Universal Robots URScript: FaiChun_9 Jan_10.script

def Machining1():
  # Default parameters:
  global speed_ms = 0.01
  global speed_rads = 0.75
  global accel_mss = 3
  global accel_radss = 1.2
  global blend_radius_m = 0.0003

  # Add subprograms here
  # Start of main program
  # Program generated by RoboDK v5.6.8 for UR10e on 10/01/2025 15:07:00
  # Using nominal kinematics.
  blend_radius_m = 0.0003
  speed_ms = 0.01
  # set_reference(p[0.340000, -0.015000, 0.001500, 0.000000, 0.000000, 0.000000])
  set_tcp(p[0.000000, 0.000000, 0.252000, 0.000000, 0.000000, 0.000000])
  # Show Tool
  movej([0.358985, -0.895332, -2.200270, -1.616787, 1.570796, 1.929781],accel_radss,speed_rads,0,blend_radius_m)
  movel([0.358985, -1.122148, -2.673539, -0.916702, 1.570796, 1.929781],accel_mss,speed_ms,0,blend_radius_m)
  #SetTool1
  #M_RunCode6
  #SetRPM60000
  speed_ms = 0.01
  #M_RunCode3
  movel([0.358985, -1.149717, -2.688845, -0.873826, 1.570796, 1.929781],accel_mss,speed_ms,0,blend_radius_m)
  speed_ms = 0.003
  movel([0.358985, -1.157003, -2.692612, -0.862774, 1.570796, 1.929781],accel_mss,speed_ms,0,blend_radius_m)
  speed_ms = 0.007
  movel([0.360284, -1.155838, -2.693115, -0.863435, 1.570796, 1.931080],accel_mss,speed_ms,0,blend_radius_m)
  movel([0.363800, -1.153166, -2.694264, -0.864959, 1.570796, 1.934596],accel_mss,speed_ms,0,blend_radius_m)
  movel([0.367667, -1.151137, -2.695132, -0.866120, 1.570796, 1.938463],accel_mss,speed_ms,0,blend_radius_m)
  movel([0.371673, -1.149666, -2.695758, -0.866965, 1.570796, 1.942469],accel_mss,speed_ms,0,blend_radius_m)
  movel([0.375593, -1.148672, -2.696180, -0.867537, 1.570796, 1.946389],accel_mss,speed_ms,0,blend_radius_m)
  movel([0.385811, -1.147094, -2.696848, -0.868447, 1.570796, 1.956607],accel_mss,speed_ms,0,blend_radius_m)
  movel([0.395233, -1.145814, -2.697388, -0.869187, 1.570796, 1.966029],accel_mss,speed_ms,0,blend_radius_m)
  movel([0.398878, -1.144990, -2.697734, -0.869664, 1.570796, 1.969674],accel_mss,speed_ms,0,blend_radius_m)
  movel([0.402533, -1.143763, -2.698250, -0.870377, 1.570796, 1.973330],accel_mss,speed_ms,0,blend_radius_m)
  movel([0.406011, -1.142059, -2.698963, -0.871368, 1.570796, 1.976808],accel_mss,speed_ms,0,blend_radius_m)
  movel([0.409148, -1.139796, -2.699904, -0.872688, 1.570796, 1.979944],accel_mss,speed_ms,0,blend_radius_m)
  movel([0.412438, -1.136413, -2.701304, -0.874672, 1.570796, 1.983234],accel_mss,speed_ms,0,blend_radius_m)
  movel([0.413570, -1.134739, -2.701992, -0.875658, 1.570796, 1.984366],accel_mss,speed_ms,0,blend_radius_m)
  movel([0.414360, -1.133075, -2.702674, -0.876641, 1.570796, 1.985156],accel_mss,speed_ms,0,blend_radius_m)
  movel([0.414991, -1.130073, -2.703896, -0.878420, 1.570796, 1.985787],accel_mss,speed_ms,0,blend_radius_m)
  movel([0.414425, -1.127699, -2.704856, -0.879834, 1.570796, 1.985221],accel_mss,speed_ms,0,blend_radius_m)
  movel([0.413477, -1.126577, -2.705309, -0.880504, 1.570796, 1.984274],accel_mss,speed_ms,0,blend_radius_m)
  movel([0.412318, -1.126143, -2.705483, -0.880763, 1.570796, 1.983114],accel_mss,speed_ms,0,blend_radius_m)
  movel([0.411061, -1.126342, -2.705403, -0.880644, 1.570796, 1.981857],accel_mss,speed_ms,0,blend_radius_m)
  movel([0.409841, -1.127103, -2.705097, -0.880189, 1.570796, 1.980638],accel_mss,speed_ms,0,blend_radius_m)
  movel([0.408484, -1.128982, -2.704338, -0.879069, 1.570796, 1.979281],accel_mss,speed_ms,0,blend_radius_m)
  movel([0.407268, -1.130867, -2.703573, -0.877948, 1.570796, 1.978064],accel_mss,speed_ms,0,blend_radius_m)
  movel([0.405338, -1.132846, -2.702767, -0.876776, 1.570796, 1.976135],accel_mss,speed_ms,0,blend_radius_m)
  movel([0.402737, -1.134615, -2.702043, -0.875731, 1.570796, 1.973533],accel_mss,speed_ms,0,blend_radius_m)
  movel([0.400364, -1.135207, -2.701800, -0.875382, 1.570796, 1.971160],accel_mss,speed_ms,0,blend_radius_m)
  movel([0.398406, -1.134766, -2.701981, -0.875642, 1.570796, 1.969202],accel_mss,speed_ms,0,blend_radius_m)
  movel([0.397035, -1.133442, -2.702523, -0.876424, 1.570796, 1.967832],accel_mss,speed_ms,0,blend_radius_m)
  movel([0.396404, -1.131466, -2.703330, -0.877593, 1.570796, 1.967200],accel_mss,speed_ms,0,blend_radius_m)
  movel([0.396662, -1.129077, -2.704300, -0.879013, 1.570796, 1.967458],accel_mss,speed_ms,0,blend_radius_m)
  movel([0.397874, -1.126522, -2.705330, -0.880536, 1.570796, 1.968671],accel_mss,speed_ms,0,blend_radius_m)
  movel([0.400111, -1.124058, -2.706319, -0.882012, 1.570796, 1.970908],accel_mss,speed_ms,0,blend_radius_m)
  movel([0.402368, -1.122361, -2.706996, -0.883031, 1.570796, 1.973164],accel_mss,speed_ms,0,blend_radius_m)
  movel([0.404592, -1.121272, -2.707430, -0.883687, 1.570796, 1.975389],accel_mss,speed_ms,0,blend_radius_m)
  movel([0.406779, -1.120798, -2.707618, -0.883973, 1.570796, 1.977575],accel_mss,speed_ms,0,blend_radius_m)
  movel([0.408920, -1.120940, -2.707561, -0.883887, 1.570796, 1.979716],accel_mss,speed_ms,0,blend_radius_m)
  movel([0.410941, -1.121627, -2.707288, -0.883473, 1.570796, 1.981737],accel_mss,speed_ms,0,blend_radius_m)
  movel([0.412761, -1.122788, -2.706826, -0.882775, 1.570796, 1.983557],accel_mss,speed_ms,0,blend_radius_m)
  movel([0.415800, -1.126514, -2.705334, -0.880541, 1.570796, 1.986596],accel_mss,speed_ms,0,blend_radius_m)
  movel([0.417144, -1.129442, -2.704152, -0.878795, 1.570796, 1.987940],accel_mss,speed_ms,0,blend_radius_m)
  movel([0.417974, -1.132572, -2.702879, -0.876938, 1.570796, 1.988771],accel_mss,speed_ms,0,blend_radius_m)
  movel([0.418302, -1.135897, -2.701516, -0.874976, 1.570796, 1.989099],accel_mss,speed_ms,0,blend_radius_m)
  movel([0.418128, -1.139411, -2.700064, -0.872914, 1.570796, 1.988924],accel_mss,speed_ms,0,blend_radius_m)
  movel([0.417267, -1.142978, -2.698578, -0.870833, 1.570796, 1.988063],accel_mss,speed_ms,0,blend_radius_m)
  movel([0.415537, -1.146458, -2.697116, -0.868815, 1.570796, 1.986334],accel_mss,speed_ms,0,blend_radius_m)
  movel([0.412946, -1.149856, -2.695677, -0.866856, 1.570796, 1.983742],accel_mss,speed_ms,0,blend_radius_m)
  movel([0.409498, -1.153176, -2.694260, -0.864954, 1.570796, 1.980294],accel_mss,speed_ms,0,blend_radius_m)
  movel([0.406063, -1.155728, -2.693163, -0.863498, 1.570796, 1.976860],accel_mss,speed_ms,0,blend_radius_m)
  movel([0.402585, -1.157607, -2.692351, -0.862431, 1.570796, 1.973381],accel_mss,speed_ms,0,blend_radius_m)
  movel([0.399151, -1.158929, -2.691777, -0.861683, 1.570796, 1.969948],accel_mss,speed_ms,0,blend_radius_m)
  movel([0.395859, -1.159805, -2.691396, -0.861188, 1.570796, 1.966655],accel_mss,speed_ms,0,blend_radius_m)
  movel([0.388031, -1.160961, -2.690892, -0.860535, 1.570796, 1.958827],accel_mss,speed_ms,0,blend_radius_m)
  movel([0.380613, -1.162143, -2.690376, -0.859870, 1.570796, 1.951410],accel_mss,speed_ms,0,blend_radius_m)
  movel([0.377615, -1.162965, -2.690015, -0.859408, 1.570796, 1.948411],accel_mss,speed_ms,0,blend_radius_m)
  movel([0.374545, -1.164177, -2.689483, -0.858729, 1.570796, 1.945341],accel_mss,speed_ms,0,blend_radius_m)
  movel([0.371509, -1.165851, -2.688746, -0.857792, 1.570796, 1.942306],accel_mss,speed_ms,0,blend_radius_m)
  movel([0.368622, -1.168057, -2.687769, -0.856563, 1.570796, 1.939418],accel_mss,speed_ms,0,blend_radius_m)
  movel([0.369262, -1.169016, -2.687343, -0.856030, 1.570796, 1.940058],accel_mss,speed_ms,0,blend_radius_m)
  movel([0.371229, -1.171492, -2.686239, -0.854659, 1.570796, 1.942025],accel_mss,speed_ms,0,blend_radius_m)
  movel([0.373363, -1.173304, -2.685426, -0.853659, 1.570796, 1.944159],accel_mss,speed_ms,0,blend_radius_m)
  movel([0.375672, -1.174449, -2.684911, -0.853029, 1.570796, 1.946468],accel_mss,speed_ms,0,blend_radius_m)
  movel([0.378153, -1.174934, -2.684692, -0.852763, 1.570796, 1.948949],accel_mss,speed_ms,0,blend_radius_m)
  movel([0.380756, -1.174836, -2.684736, -0.852816, 1.570796, 1.951553],accel_mss,speed_ms,0,blend_radius_m)
  movel([0.383422, -1.174230, -2.685010, -0.853150, 1.570796, 1.954218],accel_mss,speed_ms,0,blend_radius_m)
  movel([0.386160, -1.173110, -2.685513, -0.853766, 1.570796, 1.956957],accel_mss,speed_ms,0,blend_radius_m)
  movel([0.388972, -1.171476, -2.686246, -0.854667, 1.570796, 1.959768],accel_mss,speed_ms,0,blend_radius_m)
  movel([0.376141, -1.182465, -2.681266, -0.848658, 1.570796, 1.946938],accel_mss,speed_ms,0,blend_radius_m)
  movel([0.358985, -1.157003, -2.692612, -0.862774, 1.570796, 1.929781],accel_mss,speed_ms,0,blend_radius_m)
  speed_ms = 0.003
  movel([0.358985, -1.149717, -2.688845, -0.873826, 1.570796, 1.929781],accel_mss,speed_ms,0,blend_radius_m)
  speed_ms = 0.01
  movel([0.358985, -1.122148, -2.673539, -0.916702, 1.570796, 1.929781],accel_mss,speed_ms,0,blend_radius_m)
  #M_RunCode9
  movel([0.390070, -1.155228, -2.659313, -0.897848, 1.570796, 1.960867],accel_mss,speed_ms,0,blend_radius_m)
  #M_RunCode3
  movel([0.390070, -1.182636, -2.674188, -0.855565, 1.570796, 1.960867],accel_mss,speed_ms,0,blend_radius_m)
  speed_ms = 0.003
  movel([0.390070, -1.189858, -2.677844, -0.844687, 1.570796, 1.960867],accel_mss,speed_ms,0,blend_radius_m)
  speed_ms = 0.007
  movel([0.396700, -1.183388, -2.680842, -0.848159, 1.570796, 1.967497],accel_mss,speed_ms,0,blend_radius_m)
  movel([0.406631, -1.174785, -2.684760, -0.852845, 1.570796, 1.977428],accel_mss,speed_ms,0,blend_radius_m)
  movel([0.416940, -1.166524, -2.688448, -0.857416, 1.570796, 1.987736],accel_mss,speed_ms,0,blend_radius_m)
  movel([0.424558, -1.161153, -2.690809, -0.860427, 1.570796, 1.995354],accel_mss,speed_ms,0,blend_radius_m)
  movel([0.427380, -1.159602, -2.691485, -0.861302, 1.570796, 1.998176],accel_mss,speed_ms,0,blend_radius_m)
  movel([0.429592, -1.158857, -2.691809, -0.861723, 1.570796, 2.000389],accel_mss,speed_ms,0,blend_radius_m)
  movel([0.431192, -1.158925, -2.691779, -0.861685, 1.570796, 2.001988],accel_mss,speed_ms,0,blend_radius_m)
  movel([0.432177, -1.159797, -2.691400, -0.861192, 1.570796, 2.002973],accel_mss,speed_ms,0,blend_radius_m)
  movel([0.432434, -1.161264, -2.690760, -0.860365, 1.570796, 2.003230],accel_mss,speed_ms,0,blend_radius_m)
  movel([0.431856, -1.163109, -2.689953, -0.859328, 1.570796, 2.002653],accel_mss,speed_ms,0,blend_radius_m)
  movel([0.430453, -1.165326, -2.688977, -0.858086, 1.570796, 2.001249],accel_mss,speed_ms,0,blend_radius_m)
  movel([0.428224, -1.167916, -2.687832, -0.856641, 1.570796, 1.999021],accel_mss,speed_ms,0,blend_radius_m)
  movel([0.421358, -1.174456, -2.684908, -0.853025, 1.570796, 1.992155],accel_mss,speed_ms,0,blend_radius_m)
  movel([0.411361, -1.182965, -2.681036, -0.848388, 1.570796, 1.982158],accel_mss,speed_ms,0,blend_radius_m)
  movel([0.401263, -1.190989, -2.677315, -0.844085, 1.570796, 1.972059],accel_mss,speed_ms,0,blend_radius_m)
  movel([0.393942, -1.196149, -2.674885, -0.841355, 1.570796, 1.964739],accel_mss,speed_ms,0,blend_radius_m)
  movel([0.391243, -1.197643, -2.674176, -0.840570, 1.570796, 1.962040],accel_mss,speed_ms,0,blend_radius_m)
  movel([0.389113, -1.198381, -2.673825, -0.840183, 1.570796, 1.959910],accel_mss,speed_ms,0,blend_radius_m)
  movel([0.387547, -1.198358, -2.673836, -0.840195, 1.570796, 1.958343],accel_mss,speed_ms,0,blend_radius_m)
  movel([0.386539, -1.197580, -2.674206, -0.840603, 1.570796, 1.957335],accel_mss,speed_ms,0,blend_radius_m)
  movel([0.386213, -1.196230, -2.674847, -0.841312, 1.570796, 1.957009],accel_mss,speed_ms,0,blend_radius_m)
  movel([0.386687, -1.194496, -2.675667, -0.842226, 1.570796, 1.957483],accel_mss,speed_ms,0,blend_radius_m)
  movel([0.387972, -1.192374, -2.676665, -0.843349, 1.570796, 1.958769],accel_mss,speed_ms,0,blend_radius_m)
  movel([0.390070, -1.189858, -2.677844, -0.844687, 1.570796, 1.960867],accel_mss,speed_ms,0,blend_radius_m)
  speed_ms = 0.003
  movel([0.390070, -1.182636, -2.674188, -0.855565, 1.570796, 1.960867],accel_mss,speed_ms,0,blend_radius_m)
  speed_ms = 0.01
  movel([0.390070, -1.155228, -2.659313, -0.897848, 1.570796, 1.960867],accel_mss,speed_ms,0,blend_radius_m)
  #M_RunCode9
  movel([0.383757, -1.157911, -2.658112, -0.896367, 1.570796, 1.954554],accel_mss,speed_ms,0,blend_radius_m)
  #M_RunCode3
  movel([0.383757, -1.185302, -2.672951, -0.854136, 1.570796, 1.954554],accel_mss,speed_ms,0,blend_radius_m)
  speed_ms = 0.003
  movel([0.383757, -1.192518, -2.676598, -0.843273, 1.570796, 1.954554],accel_mss,speed_ms,0,blend_radius_m)
  speed_ms = 0.007
  movel([0.384034, -1.190067, -2.677746, -0.844576, 1.570796, 1.954830],accel_mss,speed_ms,0,blend_radius_m)
  movel([0.384719, -1.187441, -2.678969, -0.845979, 1.570796, 1.955516],accel_mss,speed_ms,0,blend_radius_m)
  movel([0.385830, -1.184674, -2.680249, -0.847465, 1.570796, 1.956626],accel_mss,speed_ms,0,blend_radius_m)
  movel([0.387369, -1.181762, -2.681588, -0.849039, 1.570796, 1.958165],accel_mss,speed_ms,0,blend_radius_m)
  movel([0.389339, -1.178702, -2.682986, -0.850702, 1.570796, 1.960136],accel_mss,speed_ms,0,blend_radius_m)
  movel([0.391735, -1.175551, -2.684414, -0.852424, 1.570796, 1.962531],accel_mss,speed_ms,0,blend_radius_m)
  movel([0.394540, -1.172369, -2.685846, -0.854174, 1.570796, 1.965337],accel_mss,speed_ms,0,blend_radius_m)
  movel([0.397760, -1.169157, -2.687280, -0.855952, 1.570796, 1.968556],accel_mss,speed_ms,0,blend_radius_m)
  movel([0.401398, -1.165917, -2.688716, -0.857755, 1.570796, 1.972194],accel_mss,speed_ms,0,blend_radius_m)
  movel([0.405183, -1.162881, -2.690052, -0.859456, 1.570796, 1.975979],accel_mss,speed_ms,0,blend_radius_m)
  movel([0.408839, -1.160283, -2.691188, -0.860918, 1.570796, 1.979636],accel_mss,speed_ms,0,blend_radius_m)
  movel([0.412361, -1.158134, -2.692122, -0.862133, 1.570796, 1.983157],accel_mss,speed_ms,0,blend_radius_m)
  movel([0.415741, -1.156438, -2.692856, -0.863094, 1.570796, 1.986537],accel_mss,speed_ms,0,blend_radius_m)
  movel([0.418920, -1.155194, -2.693393, -0.863802, 1.570796, 1.989717],accel_mss,speed_ms,0,blend_radius_m)
  movel([0.421843, -1.154407, -2.693731, -0.864250, 1.570796, 1.992639],accel_mss,speed_ms,0,blend_radius_m)
  movel([0.424499, -1.154076, -2.693874, -0.864439, 1.570796, 1.995295],accel_mss,speed_ms,0,blend_radius_m)
  movel([0.426890, -1.154203, -2.693819, -0.864367, 1.570796, 1.997687],accel_mss,speed_ms,0,blend_radius_m)
  movel([0.428991, -1.154756, -2.693581, -0.864051, 1.570796, 1.999787],accel_mss,speed_ms,0,blend_radius_m)
  movel([0.430782, -1.155707, -2.693172, -0.863511, 1.570796, 2.001578],accel_mss,speed_ms,0,blend_radius_m)
  movel([0.432260, -1.157045, -2.692594, -0.862750, 1.570796, 2.003056],accel_mss,speed_ms,0,blend_radius_m)
  movel([0.433430, -1.158771, -2.691846, -0.861772, 1.570796, 2.004226],accel_mss,speed_ms,0,blend_radius_m)
  movel([0.434237, -1.160788, -2.690968, -0.860633, 1.570796, 2.005033],accel_mss,speed_ms,0,blend_radius_m)
  movel([0.434638, -1.162993, -2.690003, -0.859393, 1.570796, 2.005434],accel_mss,speed_ms,0,blend_radius_m)
  movel([0.434635, -1.165385, -2.688951, -0.858052, 1.570796, 2.005431],accel_mss,speed_ms,0,blend_radius_m)
  movel([0.434233, -1.167961, -2.687812, -0.856616, 1.570796, 2.005030],accel_mss,speed_ms,0,blend_radius_m)
  movel([0.433415, -1.170685, -2.686599, -0.855105, 1.570796, 2.004211],accel_mss,speed_ms,0,blend_radius_m)
  movel([0.432178, -1.173518, -2.685330, -0.853541, 1.570796, 2.002974],accel_mss,speed_ms,0,blend_radius_m)
  movel([0.430522, -1.176455, -2.684005, -0.851929, 1.570796, 2.001318],accel_mss,speed_ms,0,blend_radius_m)
  movel([0.428448, -1.179502, -2.682621, -0.850266, 1.570796, 1.999245],accel_mss,speed_ms,0,blend_radius_m)
  movel([0.425982, -1.182592, -2.681208, -0.848589, 1.570796, 1.996779],accel_mss,speed_ms,0,blend_radius_m)
  movel([0.423147, -1.185664, -2.679792, -0.846933, 1.570796, 1.993943],accel_mss,speed_ms,0,blend_radius_m)
  movel([0.419941, -1.188728, -2.678370, -0.845290, 1.570796, 1.990737],accel_mss,speed_ms,0,blend_radius_m)
  movel([0.416367, -1.191779, -2.676945, -0.843665, 1.570796, 1.987163],accel_mss,speed_ms,0,blend_radius_m)
  movel([0.412690, -1.194608, -2.675614, -0.842167, 1.570796, 1.983486],accel_mss,speed_ms,0,blend_radius_m)
  movel([0.409169, -1.197005, -2.674479, -0.840905, 1.570796, 1.979965],accel_mss,speed_ms,0,blend_radius_m)
  movel([0.405805, -1.198977, -2.673541, -0.839871, 1.570796, 1.976601],accel_mss,speed_ms,0,blend_radius_m)
  movel([0.402584, -1.200530, -2.672799, -0.839060, 1.570796, 1.973380],accel_mss,speed_ms,0,blend_radius_m)
  movel([0.399556, -1.201668, -2.672254, -0.838467, 1.570796, 1.970353],accel_mss,speed_ms,0,blend_radius_m)
  movel([0.396767, -1.202400, -2.671902, -0.838087, 1.570796, 1.967564],accel_mss,speed_ms,0,blend_radius_m)
  movel([0.394210, -1.202727, -2.671745, -0.837916, 1.570796, 1.965007],accel_mss,speed_ms,0,blend_radius_m)
  movel([0.391887, -1.202647, -2.671784, -0.837958, 1.570796, 1.962683],accel_mss,speed_ms,0,blend_radius_m)
  movel([0.389820, -1.202186, -2.672006, -0.838198, 1.570796, 1.960616],accel_mss,speed_ms,0,blend_radius_m)
  movel([0.388028, -1.201364, -2.672400, -0.838625, 1.570796, 1.958824],accel_mss,speed_ms,0,blend_radius_m)
  movel([0.386519, -1.200177, -2.672968, -0.839244, 1.570796, 1.957315],accel_mss,speed_ms,0,blend_radius_m)
  movel([0.385286, -1.198629, -2.673707, -0.840053, 1.570796, 1.956082],accel_mss,speed_ms,0,blend_radius_m)
  movel([0.384388, -1.196795, -2.674579, -0.841015, 1.570796, 1.955184],accel_mss,speed_ms,0,blend_radius_m)
  movel([0.383876, -1.194758, -2.675543, -0.842088, 1.570796, 1.954672],accel_mss,speed_ms,0,blend_radius_m)
  movel([0.383757, -1.192518, -2.676598, -0.843273, 1.570796, 1.954554],accel_mss,speed_ms,0,blend_radius_m)
  speed_ms = 0.003
  movel([0.383757, -1.185302, -2.672951, -0.854136, 1.570796, 1.954554],accel_mss,speed_ms,0,blend_radius_m)
  speed_ms = 0.01
  movel([0.383757, -1.157911, -2.658112, -0.896367, 1.570796, 1.954554],accel_mss,speed_ms,0,blend_radius_m)
  #M_RunCode9
  movel([0.496093, -1.382466, -2.528375, -0.801548, 1.570796, 2.066889],accel_mss,speed_ms,0,blend_radius_m)
  #M_RunCode3
  movel([0.496093, -1.406789, -2.540293, -0.765307, 1.570796, 2.066889],accel_mss,speed_ms,0,blend_radius_m)
  speed_ms = 0.003
  movel([0.496093, -1.413093, -2.543201, -0.756095, 1.570796, 2.066889],accel_mss,speed_ms,0,blend_radius_m)
  speed_ms = 0.007
  movel([0.497104, -1.412495, -2.543652, -0.756242, 1.570796, 2.067901],accel_mss,speed_ms,0,blend_radius_m)
  movel([0.499783, -1.411227, -2.544607, -0.756556, 1.570796, 2.070579],accel_mss,speed_ms,0,blend_radius_m)
  movel([0.502622, -1.410494, -2.545157, -0.756738, 1.570796, 2.073418],accel_mss,speed_ms,0,blend_radius_m)
  movel([0.505487, -1.410196, -2.545381, -0.756812, 1.570796, 2.076283],accel_mss,speed_ms,0,blend_radius_m)
  movel([0.508237, -1.410226, -2.545358, -0.756805, 1.570796, 2.079034],accel_mss,speed_ms,0,blend_radius_m)
  movel([0.515289, -1.411028, -2.544756, -0.756605, 1.570796, 2.086086],accel_mss,speed_ms,0,blend_radius_m)
  movel([0.521765, -1.411881, -2.544115, -0.756394, 1.570796, 2.092561],accel_mss,speed_ms,0,blend_radius_m)
  movel([0.524304, -1.411969, -2.544048, -0.756372, 1.570796, 2.095101],accel_mss,speed_ms,0,blend_radius_m)
  movel([0.526887, -1.411770, -2.544198, -0.756421, 1.570796, 2.097684],accel_mss,speed_ms,0,blend_radius_m)
  movel([0.529402, -1.411199, -2.544627, -0.756563, 1.570796, 2.100198],accel_mss,speed_ms,0,blend_radius_m)
  movel([0.531734, -1.410169, -2.545401, -0.756819, 1.570796, 2.102530],accel_mss,speed_ms,0,blend_radius_m)
  movel([0.534284, -1.408370, -2.546748, -0.757271, 1.570796, 2.105081],accel_mss,speed_ms,0,blend_radius_m)
  movel([0.535210, -1.407391, -2.547480, -0.757519, 1.570796, 2.106007],accel_mss,speed_ms,0,blend_radius_m)
  movel([0.535902, -1.406358, -2.548250, -0.757782, 1.570796, 2.106698],accel_mss,speed_ms,0,blend_radius_m)
  movel([0.536626, -1.404345, -2.549745, -0.758299, 1.570796, 2.107423],accel_mss,speed_ms,0,blend_radius_m)
  movel([0.536483, -1.402557, -2.551069, -0.758763, 1.570796, 2.107279],accel_mss,speed_ms,0,blend_radius_m)
  movel([0.535964, -1.401585, -2.551787, -0.759017, 1.570796, 2.106761],accel_mss,speed_ms,0,blend_radius_m)
  movel([0.535230, -1.401062, -2.552172, -0.759155, 1.570796, 2.106027],accel_mss,speed_ms,0,blend_radius_m)
  movel([0.534373, -1.400967, -2.552242, -0.759180, 1.570796, 2.105170],accel_mss,speed_ms,0,blend_radius_m)
  movel([0.533483, -1.401277, -2.552014, -0.759098, 1.570796, 2.104279],accel_mss,speed_ms,0,blend_radius_m)
  movel([0.532384, -1.402355, -2.551218, -0.758816, 1.570796, 2.103180],accel_mss,speed_ms,0,blend_radius_m)
  movel([0.531379, -1.403465, -2.550397, -0.758527, 1.570796, 2.102176],accel_mss,speed_ms,0,blend_radius_m)
  movel([0.529890, -1.404508, -2.549624, -0.758257, 1.570796, 2.100686],accel_mss,speed_ms,0,blend_radius_m)
  movel([0.527963, -1.405280, -2.549051, -0.758058, 1.570796, 2.098760],accel_mss,speed_ms,0,blend_radius_m)
  movel([0.526316, -1.405254, -2.549070, -0.758064, 1.570796, 2.097112],accel_mss,speed_ms,0,blend_radius_m)
  movel([0.525050, -1.404571, -2.549577, -0.758240, 1.570796, 2.095846],accel_mss,speed_ms,0,blend_radius_m)
  movel([0.524270, -1.403366, -2.550470, -0.758552, 1.570796, 2.095067],accel_mss,speed_ms,0,blend_radius_m)
  movel([0.524055, -1.401836, -2.551601, -0.758951, 1.570796, 2.094851],accel_mss,speed_ms,0,blend_radius_m)
  movel([0.524478, -1.400181, -2.552821, -0.759387, 1.570796, 2.095274],accel_mss,speed_ms,0,blend_radius_m)
  movel([0.525555, -1.398592, -2.553988, -0.759809, 1.570796, 2.096352],accel_mss,speed_ms,0,blend_radius_m)
  movel([0.527302, -1.397266, -2.554959, -0.760164, 1.570796, 2.098099],accel_mss,speed_ms,0,blend_radius_m)
  movel([0.528984, -1.396492, -2.555524, -0.760372, 1.570796, 2.099781],accel_mss,speed_ms,0,blend_radius_m)
  movel([0.530578, -1.396145, -2.555778, -0.760466, 1.570796, 2.101374],accel_mss,speed_ms,0,blend_radius_m)
  movel([0.532081, -1.396224, -2.555720, -0.760445, 1.570796, 2.102877],accel_mss,speed_ms,0,blend_radius_m)
  movel([0.533493, -1.396734, -2.555347, -0.760307, 1.570796, 2.104290],accel_mss,speed_ms,0,blend_radius_m)
  movel([0.534769, -1.397605, -2.554711, -0.760073, 1.570796, 2.105566],accel_mss,speed_ms,0,blend_radius_m)
  movel([0.535865, -1.398770, -2.553857, -0.759762, 1.570796, 2.106661],accel_mss,speed_ms,0,blend_radius_m)
  movel([0.537521, -1.401976, -2.551498, -0.758915, 1.570796, 2.108317],accel_mss,speed_ms,0,blend_radius_m)
  movel([0.538126, -1.404299, -2.549779, -0.758311, 1.570796, 2.108923],accel_mss,speed_ms,0,blend_radius_m)
  movel([0.538374, -1.406672, -2.548015, -0.757702, 1.570796, 2.109170],accel_mss,speed_ms,0,blend_radius_m)
  movel([0.538264, -1.409089, -2.546211, -0.757090, 1.570796, 2.109060],accel_mss,speed_ms,0,blend_radius_m)
  movel([0.537801, -1.411550, -2.544364, -0.756476, 1.570796, 2.108597],accel_mss,speed_ms,0,blend_radius_m)
  movel([0.536875, -1.413924, -2.542573, -0.755892, 1.570796, 2.107671],accel_mss,speed_ms,0,blend_radius_m)
  movel([0.535368, -1.416086, -2.540936, -0.755367, 1.570796, 2.106164],accel_mss,speed_ms,0,blend_radius_m)
  movel([0.533284, -1.418039, -2.539451, -0.754899, 1.570796, 2.104080],accel_mss,speed_ms,0,blend_radius_m)
  movel([0.530625, -1.419784, -2.538119, -0.754486, 1.570796, 2.101421],accel_mss,speed_ms,0,blend_radius_m)
  movel([0.528047, -1.420988, -2.537198, -0.754204, 1.570796, 2.098844],accel_mss,speed_ms,0,blend_radius_m)
  movel([0.525504, -1.421702, -2.536650, -0.754037, 1.570796, 2.096300],accel_mss,speed_ms,0,blend_radius_m)
  movel([0.523046, -1.422024, -2.536403, -0.753962, 1.570796, 2.093842],accel_mss,speed_ms,0,blend_radius_m)
  movel([0.520727, -1.422052, -2.536382, -0.753956, 1.570796, 2.091523],accel_mss,speed_ms,0,blend_radius_m)
  movel([0.515303, -1.421445, -2.536847, -0.754097, 1.570796, 2.086099],accel_mss,speed_ms,0,blend_radius_m)
  movel([0.510152, -1.420924, -2.537247, -0.754219, 1.570796, 2.080948],accel_mss,speed_ms,0,blend_radius_m)
  movel([0.508029, -1.420964, -2.537216, -0.754209, 1.570796, 2.078825],accel_mss,speed_ms,0,blend_radius_m)
  movel([0.505817, -1.421270, -2.536982, -0.754138, 1.570796, 2.076613],accel_mss,speed_ms,0,blend_radius_m)
  movel([0.503574, -1.421917, -2.536485, -0.753987, 1.570796, 2.074370],accel_mss,speed_ms,0,blend_radius_m)
  movel([0.501367, -1.422986, -2.535664, -0.753740, 1.570796, 2.072163],accel_mss,speed_ms,0,blend_radius_m)
  movel([0.501695, -1.423803, -2.535035, -0.753552, 1.570796, 2.072492],accel_mss,speed_ms,0,blend_radius_m)
  movel([0.502756, -1.425977, -2.533355, -0.753056, 1.570796, 2.073552],accel_mss,speed_ms,0,blend_radius_m)
  movel([0.504008, -1.427693, -2.532026, -0.752670, 1.570796, 2.074805],accel_mss,speed_ms,0,blend_radius_m)
  movel([0.505454, -1.428956, -2.531044, -0.752389, 1.570796, 2.076250],accel_mss,speed_ms,0,blend_radius_m)
  movel([0.507091, -1.429766, -2.530413, -0.752210, 1.570796, 2.077887],accel_mss,speed_ms,0,blend_radius_m)
  movel([0.508876, -1.430170, -2.530098, -0.752121, 1.570796, 2.079672],accel_mss,speed_ms,0,blend_radius_m)
  movel([0.510757, -1.430216, -2.530063, -0.752111, 1.570796, 2.081553],accel_mss,speed_ms,0,blend_radius_m)
  movel([0.512740, -1.429904, -2.530306, -0.752179, 1.570796, 2.083536],accel_mss,speed_ms,0,blend_radius_m)
  movel([0.514827, -1.429230, -2.530831, -0.752328, 1.570796, 2.085623],accel_mss,speed_ms,0,blend_radius_m)
  movel([0.504898, -1.434894, -2.526397, -0.751098, 1.570796, 2.075694],accel_mss,speed_ms,0,blend_radius_m)
  movel([0.496093, -1.413093, -2.543201, -0.756095, 1.570796, 2.066889],accel_mss,speed_ms,0,blend_radius_m)
  speed_ms = 0.003
  movel([0.496093, -1.406789, -2.540293, -0.765307, 1.570796, 2.066889],accel_mss,speed_ms,0,blend_radius_m)
  speed_ms = 0.01
  movel([0.496093, -1.382466, -2.528375, -0.801548, 1.570796, 2.066889],accel_mss,speed_ms,0,blend_radius_m)
  #M_RunCode9
  movel([0.512138, -1.403973, -2.512554, -0.795862, 1.570796, 2.082934],accel_mss,speed_ms,0,blend_radius_m)
  #M_RunCode3
  movel([0.512138, -1.427879, -2.524206, -0.760304, 1.570796, 2.082934],accel_mss,speed_ms,0,blend_radius_m)
  speed_ms = 0.003
  movel([0.512138, -1.434068, -2.527046, -0.751275, 1.570796, 2.082934],accel_mss,speed_ms,0,blend_radius_m)
  speed_ms = 0.007
  movel([0.514003, -1.433320, -2.527634, -0.751435, 1.570796, 2.084799],accel_mss,speed_ms,0,blend_radius_m)
  movel([0.515626, -1.433332, -2.527624, -0.751432, 1.570796, 2.086422],accel_mss,speed_ms,0,blend_radius_m)
  movel([0.516887, -1.433975, -2.527119, -0.751294, 1.570796, 2.087684],accel_mss,speed_ms,0,blend_radius_m)
  movel([0.517657, -1.435128, -2.526212, -0.751048, 1.570796, 2.088453],accel_mss,speed_ms,0,blend_radius_m)
  movel([0.517868, -1.436594, -2.525056, -0.750738, 1.570796, 2.088665],accel_mss,speed_ms,0,blend_radius_m)
  movel([0.517453, -1.438175, -2.523806, -0.750408, 1.570796, 2.088249],accel_mss,speed_ms,0,blend_radius_m)
  movel([0.516413, -1.439679, -2.522613, -0.750097, 1.570796, 2.087209],accel_mss,speed_ms,0,blend_radius_m)
  movel([0.514754, -1.440917, -2.521629, -0.749844, 1.570796, 2.085550],accel_mss,speed_ms,0,blend_radius_m)
  movel([0.513217, -1.441589, -2.521093, -0.749707, 1.570796, 2.084014],accel_mss,speed_ms,0,blend_radius_m)
  movel([0.511950, -1.441787, -2.520935, -0.749667, 1.570796, 2.082746],accel_mss,speed_ms,0,blend_radius_m)
  movel([0.510647, -1.442088, -2.520695, -0.749606, 1.570796, 2.081443],accel_mss,speed_ms,0,blend_radius_m)
  movel([0.509919, -1.442689, -2.520215, -0.749485, 1.570796, 2.080715],accel_mss,speed_ms,0,blend_radius_m)
  movel([0.509449, -1.443526, -2.519546, -0.749317, 1.570796, 2.080245],accel_mss,speed_ms,0,blend_radius_m)
  movel([0.509278, -1.444452, -2.518804, -0.749133, 1.570796, 2.080074],accel_mss,speed_ms,0,blend_radius_m)
  movel([0.509440, -1.445324, -2.518105, -0.748960, 1.570796, 2.080236],accel_mss,speed_ms,0,blend_radius_m)
  movel([0.509993, -1.446284, -2.517333, -0.748772, 1.570796, 2.080789],accel_mss,speed_ms,0,blend_radius_m)
  movel([0.510801, -1.446988, -2.516767, -0.748634, 1.570796, 2.081597],accel_mss,speed_ms,0,blend_radius_m)
  movel([0.511865, -1.447436, -2.516405, -0.748547, 1.570796, 2.082661],accel_mss,speed_ms,0,blend_radius_m)
  movel([0.513186, -1.447631, -2.516249, -0.748510, 1.570796, 2.083982],accel_mss,speed_ms,0,blend_radius_m)
  movel([0.514688, -1.447559, -2.516306, -0.748524, 1.570796, 2.085484],accel_mss,speed_ms,0,blend_radius_m)
  movel([0.516291, -1.447213, -2.516585, -0.748591, 1.570796, 2.087087],accel_mss,speed_ms,0,blend_radius_m)
  movel([0.517999, -1.446591, -2.517086, -0.748712, 1.570796, 2.088795],accel_mss,speed_ms,0,blend_radius_m)
  movel([0.519813, -1.445693, -2.517809, -0.748888, 1.570796, 2.090609],accel_mss,speed_ms,0,blend_radius_m)
  movel([0.522666, -1.443719, -2.519391, -0.749279, 1.570796, 2.093462],accel_mss,speed_ms,0,blend_radius_m)
  movel([0.524983, -1.441258, -2.521357, -0.749774, 1.570796, 2.095780],accel_mss,speed_ms,0,blend_radius_m)
  movel([0.525915, -1.439851, -2.522477, -0.750062, 1.570796, 2.096711],accel_mss,speed_ms,0,blend_radius_m)
  movel([0.526652, -1.438341, -2.523675, -0.750373, 1.570796, 2.097449],accel_mss,speed_ms,0,blend_radius_m)
  movel([0.527554, -1.435008, -2.526307, -0.751074, 1.570796, 2.098351],accel_mss,speed_ms,0,blend_radius_m)
  movel([0.527587, -1.431347, -2.529179, -0.751863, 1.570796, 2.098383],accel_mss,speed_ms,0,blend_radius_m)
  movel([0.526637, -1.427456, -2.532210, -0.752723, 1.570796, 2.097433],accel_mss,speed_ms,0,blend_radius_m)
  movel([0.542111, -1.418898, -2.538796, -0.754695, 1.570796, 2.112907],accel_mss,speed_ms,0,blend_radius_m)
  movel([0.547688, -1.435758, -2.525716, -0.750915, 1.570796, 2.118485],accel_mss,speed_ms,0,blend_radius_m)
  movel([0.537746, -1.441111, -2.521474, -0.749804, 1.570796, 2.108543],accel_mss,speed_ms,0,blend_radius_m)
  movel([0.539901, -1.439199, -2.522994, -0.750196, 1.570796, 2.110697],accel_mss,speed_ms,0,blend_radius_m)
  movel([0.541670, -1.436872, -2.524837, -0.750680, 1.570796, 2.112466],accel_mss,speed_ms,0,blend_radius_m)
  movel([0.542959, -1.434240, -2.526912, -0.751238, 1.570796, 2.113756],accel_mss,speed_ms,0,blend_radius_m)
  movel([0.543680, -1.431418, -2.529124, -0.751847, 1.570796, 2.114477],accel_mss,speed_ms,0,blend_radius_m)
  movel([0.543769, -1.428514, -2.531388, -0.752487, 1.570796, 2.114565],accel_mss,speed_ms,0,blend_radius_m)
  movel([0.543166, -1.425645, -2.533613, -0.753131, 1.570796, 2.113962],accel_mss,speed_ms,0,blend_radius_m)
  movel([0.531802, -1.431868, -2.528772, -0.751749, 1.570796, 2.102598],accel_mss,speed_ms,0,blend_radius_m)
  movel([0.532645, -1.435321, -2.526060, -0.751007, 1.570796, 2.103441],accel_mss,speed_ms,0,blend_radius_m)
  movel([0.532812, -1.438966, -2.523179, -0.750244, 1.570796, 2.103608],accel_mss,speed_ms,0,blend_radius_m)
  movel([0.532201, -1.442603, -2.520284, -0.749502, 1.570796, 2.102997],accel_mss,speed_ms,0,blend_radius_m)
  movel([0.531565, -1.444346, -2.518889, -0.749154, 1.570796, 2.102361],accel_mss,speed_ms,0,blend_radius_m)
  movel([0.530709, -1.446043, -2.517527, -0.748819, 1.570796, 2.101506],accel_mss,speed_ms,0,blend_radius_m)
  movel([0.529618, -1.447639, -2.516242, -0.748508, 1.570796, 2.100414],accel_mss,speed_ms,0,blend_radius_m)
  movel([0.528273, -1.449088, -2.515072, -0.748229, 1.570796, 2.099070],accel_mss,speed_ms,0,blend_radius_m)
  movel([0.526675, -1.450389, -2.514018, -0.747982, 1.570796, 2.097472],accel_mss,speed_ms,0,blend_radius_m)
  movel([0.524823, -1.451546, -2.513080, -0.747764, 1.570796, 2.095619],accel_mss,speed_ms,0,blend_radius_m)
  movel([0.522889, -1.452474, -2.512325, -0.747590, 1.570796, 2.093685],accel_mss,speed_ms,0,blend_radius_m)
  movel([0.521038, -1.453096, -2.511818, -0.747475, 1.570796, 2.091834],accel_mss,speed_ms,0,blend_radius_m)
  movel([0.519270, -1.453408, -2.511564, -0.747417, 1.570796, 2.090067],accel_mss,speed_ms,0,blend_radius_m)
  movel([0.517584, -1.453415, -2.511558, -0.747416, 1.570796, 2.088380],accel_mss,speed_ms,0,blend_radius_m)
  movel([0.514548, -1.452701, -2.512140, -0.747548, 1.570796, 2.085344],accel_mss,speed_ms,0,blend_radius_m)
  movel([0.512020, -1.451143, -2.513407, -0.747839, 1.570796, 2.082816],accel_mss,speed_ms,0,blend_radius_m)
  movel([0.510039, -1.448945, -2.515187, -0.748257, 1.570796, 2.080835],accel_mss,speed_ms,0,blend_radius_m)
  movel([0.508638, -1.446319, -2.517305, -0.748765, 1.570796, 2.079434],accel_mss,speed_ms,0,blend_radius_m)
  movel([0.508085, -1.444283, -2.518939, -0.749166, 1.570796, 2.078881],accel_mss,speed_ms,0,blend_radius_m)
  movel([0.507919, -1.441997, -2.520768, -0.749624, 1.570796, 2.078716],accel_mss,speed_ms,0,blend_radius_m)
  movel([0.508199, -1.439645, -2.522640, -0.750104, 1.570796, 2.078995],accel_mss,speed_ms,0,blend_radius_m)
  movel([0.508988, -1.437423, -2.524402, -0.750565, 1.570796, 2.079784],accel_mss,speed_ms,0,blend_radius_m)
  movel([0.510296, -1.435505, -2.525915, -0.750968, 1.570796, 2.081093],accel_mss,speed_ms,0,blend_radius_m)
  movel([0.512138, -1.434068, -2.527046, -0.751275, 1.570796, 2.082934],accel_mss,speed_ms,0,blend_radius_m)
  speed_ms = 0.003
  movel([0.512138, -1.427879, -2.524206, -0.760304, 1.570796, 2.082934],accel_mss,speed_ms,0,blend_radius_m)
  speed_ms = 0.01
  movel([0.512138, -1.403973, -2.512554, -0.795862, 1.570796, 2.082934],accel_mss,speed_ms,0,blend_radius_m)
  #M_RunCode9
  movel([0.519767, -1.313113, -2.575087, -0.824188, 1.570796, 2.090564],accel_mss,speed_ms,0,blend_radius_m)
  #M_RunCode3
  movel([0.519767, -1.338670, -2.587888, -0.785832, 1.570796, 2.090564],accel_mss,speed_ms,0,blend_radius_m)
  speed_ms = 0.003
  movel([0.519767, -1.345323, -2.591017, -0.776049, 1.570796, 2.090564],accel_mss,speed_ms,0,blend_radius_m)
  speed_ms = 0.007
  movel([0.516626, -1.345909, -2.590631, -0.775849, 1.570796, 2.087422],accel_mss,speed_ms,0,blend_radius_m)
  movel([0.513583, -1.345852, -2.590668, -0.775868, 1.570796, 2.084379],accel_mss,speed_ms,0,blend_radius_m)
  movel([0.510695, -1.345269, -2.591053, -0.776068, 1.570796, 2.081491],accel_mss,speed_ms,0,blend_radius_m)
  movel([0.508037, -1.344256, -2.591718, -0.776415, 1.570796, 2.078833],accel_mss,speed_ms,0,blend_radius_m)
  movel([0.505666, -1.342928, -2.592588, -0.776873, 1.570796, 2.076462],accel_mss,speed_ms,0,blend_radius_m)
  movel([0.507474, -1.339287, -2.594962, -0.778140, 1.570796, 2.078270],accel_mss,speed_ms,0,blend_radius_m)
  movel([0.510328, -1.335396, -2.597479, -0.779514, 1.570796, 2.081124],accel_mss,speed_ms,0,blend_radius_m)
  movel([0.513928, -1.331601, -2.599914, -0.780873, 1.570796, 2.084724],accel_mss,speed_ms,0,blend_radius_m)
  movel([0.517969, -1.328267, -2.602038, -0.782084, 1.570796, 2.088765],accel_mss,speed_ms,0,blend_radius_m)
  movel([0.522131, -1.325765, -2.603621, -0.783002, 1.570796, 2.092928],accel_mss,speed_ms,0,blend_radius_m)
  movel([0.524156, -1.324940, -2.604142, -0.783307, 1.570796, 2.094953],accel_mss,speed_ms,0,blend_radius_m)
  movel([0.526089, -1.324461, -2.604443, -0.783485, 1.570796, 2.096885],accel_mss,speed_ms,0,blend_radius_m)
  movel([0.527884, -1.324376, -2.604497, -0.783516, 1.570796, 2.098680],accel_mss,speed_ms,0,blend_radius_m)
  movel([0.529506, -1.324725, -2.604277, -0.783387, 1.570796, 2.100302],accel_mss,speed_ms,0,blend_radius_m)
  movel([0.530909, -1.325555, -2.603754, -0.783080, 1.570796, 2.101705],accel_mss,speed_ms,0,blend_radius_m)
  movel([0.532052, -1.326908, -2.602899, -0.782582, 1.570796, 2.102848],accel_mss,speed_ms,0,blend_radius_m)
  movel([0.532898, -1.329482, -2.601266, -0.781641, 1.570796, 2.103694],accel_mss,speed_ms,0,blend_radius_m)
  movel([0.532604, -1.332369, -2.599423, -0.780597, 1.570796, 2.103400],accel_mss,speed_ms,0,blend_radius_m)
  movel([0.531317, -1.335443, -2.597449, -0.779497, 1.570796, 2.102113],accel_mss,speed_ms,0,blend_radius_m)
  movel([0.529167, -1.338587, -2.595416, -0.778385, 1.570796, 2.099963],accel_mss,speed_ms,0,blend_radius_m)
  movel([0.526095, -1.341783, -2.593337, -0.777269, 1.570796, 2.096891],accel_mss,speed_ms,0,blend_radius_m)
  movel([0.522942, -1.343988, -2.591894, -0.776507, 1.570796, 2.093738],accel_mss,speed_ms,0,blend_radius_m)
  movel([0.519767, -1.345323, -2.591017, -0.776049, 1.570796, 2.090564],accel_mss,speed_ms,0,blend_radius_m)
  speed_ms = 0.003
  movel([0.519767, -1.338670, -2.587888, -0.785832, 1.570796, 2.090564],accel_mss,speed_ms,0,blend_radius_m)
  speed_ms = 0.01
  movel([0.519767, -1.313113, -2.575087, -0.824188, 1.570796, 2.090564],accel_mss,speed_ms,0,blend_radius_m)
  #M_RunCode9
  movel([0.614162, -1.215204, -2.630657, -0.866528, 1.570796, 2.184958],accel_mss,speed_ms,0,blend_radius_m)
  #M_RunCode3
  movel([0.614162, -1.242100, -2.644742, -0.825547, 1.570796, 2.184958],accel_mss,speed_ms,0,blend_radius_m)
  speed_ms = 0.003
  movel([0.614162, -1.249153, -2.648196, -0.815040, 1.570796, 2.184958],accel_mss,speed_ms,0,blend_radius_m)
  speed_ms = 0.007
  movel([0.612984, -1.247832, -2.648901, -0.815656, 1.570796, 2.183781],accel_mss,speed_ms,0,blend_radius_m)
  movel([0.612328, -1.246039, -2.649854, -0.816496, 1.570796, 2.183124],accel_mss,speed_ms,0,blend_radius_m)
  movel([0.611967, -1.244003, -2.650932, -0.817454, 1.570796, 2.182763],accel_mss,speed_ms,0,blend_radius_m)
  movel([0.612891, -1.243759, -2.651061, -0.817569, 1.570796, 2.183688],accel_mss,speed_ms,0,blend_radius_m)
  movel([0.613408, -1.244165, -2.650846, -0.817377, 1.570796, 2.184205],accel_mss,speed_ms,0,blend_radius_m)
  movel([0.614057, -1.244575, -2.650629, -0.817184, 1.570796, 2.184853],accel_mss,speed_ms,0,blend_radius_m)
  movel([0.615382, -1.244348, -2.650750, -0.817291, 1.570796, 2.186178],accel_mss,speed_ms,0,blend_radius_m)
  movel([0.616875, -1.243518, -2.651188, -0.817683, 1.570796, 2.187672],accel_mss,speed_ms,0,blend_radius_m)
  movel([0.618326, -1.242417, -2.651768, -0.818204, 1.570796, 2.189123],accel_mss,speed_ms,0,blend_radius_m)
  movel([0.620313, -1.240830, -2.652602, -0.818957, 1.570796, 2.191110],accel_mss,speed_ms,0,blend_radius_m)
  movel([0.620034, -1.238169, -2.653993, -0.820227, 1.570796, 2.190831],accel_mss,speed_ms,0,blend_radius_m)
  movel([0.619026, -1.236416, -2.654905, -0.821068, 1.570796, 2.189822],accel_mss,speed_ms,0,blend_radius_m)
  movel([0.618176, -1.236010, -2.655115, -0.821263, 1.570796, 2.188973],accel_mss,speed_ms,0,blend_radius_m)
  movel([0.617059, -1.235990, -2.655126, -0.821273, 1.570796, 2.187855],accel_mss,speed_ms,0,blend_radius_m)
  movel([0.615652, -1.236407, -2.654910, -0.821072, 1.570796, 2.186449],accel_mss,speed_ms,0,blend_radius_m)
  movel([0.613924, -1.237313, -2.654439, -0.820638, 1.570796, 2.184720],accel_mss,speed_ms,0,blend_radius_m)
  movel([0.614647, -1.235492, -2.655384, -0.821513, 1.570796, 2.185444],accel_mss,speed_ms,0,blend_radius_m)
  movel([0.615472, -1.233933, -2.656191, -0.822266, 1.570796, 2.186268],accel_mss,speed_ms,0,blend_radius_m)
  movel([0.615964, -1.233385, -2.656473, -0.822531, 1.570796, 2.186760],accel_mss,speed_ms,0,blend_radius_m)
  movel([0.616530, -1.233065, -2.656638, -0.822686, 1.570796, 2.187326],accel_mss,speed_ms,0,blend_radius_m)
  movel([0.617945, -1.233326, -2.656504, -0.822559, 1.570796, 2.188742],accel_mss,speed_ms,0,blend_radius_m)
  movel([0.620016, -1.235079, -2.655598, -0.821712, 1.570796, 2.190813],accel_mss,speed_ms,0,blend_radius_m)
  movel([0.621390, -1.237540, -2.654321, -0.820529, 1.570796, 2.192187],accel_mss,speed_ms,0,blend_radius_m)
  movel([0.621652, -1.238983, -2.653568, -0.819838, 1.570796, 2.192448],accel_mss,speed_ms,0,blend_radius_m)
  movel([0.621543, -1.240537, -2.652755, -0.819097, 1.570796, 2.192339],accel_mss,speed_ms,0,blend_radius_m)
  movel([0.620996, -1.242179, -2.651893, -0.818317, 1.570796, 2.191793],accel_mss,speed_ms,0,blend_radius_m)
  movel([0.619955, -1.243886, -2.650993, -0.817509, 1.570796, 2.190751],accel_mss,speed_ms,0,blend_radius_m)
  movel([0.618594, -1.242857, -2.651536, -0.817995, 1.570796, 2.189390],accel_mss,speed_ms,0,blend_radius_m)
  movel([0.616086, -1.249771, -2.647866, -0.814752, 1.570796, 2.186882],accel_mss,speed_ms,0,blend_radius_m)
  movel([0.614162, -1.249153, -2.648196, -0.815040, 1.570796, 2.184958],accel_mss,speed_ms,0,blend_radius_m)
  speed_ms = 0.003
  movel([0.614162, -1.242100, -2.644742, -0.825547, 1.570796, 2.184958],accel_mss,speed_ms,0,blend_radius_m)
  speed_ms = 0.01
  movel([0.614162, -1.215204, -2.630657, -0.866528, 1.570796, 2.184958],accel_mss,speed_ms,0,blend_radius_m)
  #M_RunCode9
  movel([0.593907, -1.167128, -2.653928, -0.891333, 1.570796, 2.164704],accel_mss,speed_ms,0,blend_radius_m)
  #M_RunCode3
  movel([0.593907, -1.194457, -2.668646, -0.849286, 1.570796, 2.164704],accel_mss,speed_ms,0,blend_radius_m)
  speed_ms = 0.003
  movel([0.593907, -1.201650, -2.672262, -0.838476, 1.570796, 2.164704],accel_mss,speed_ms,0,blend_radius_m)
  speed_ms = 0.007
  movel([0.590839, -1.203902, -2.671179, -0.837308, 1.570796, 2.161636],accel_mss,speed_ms,0,blend_radius_m)
  movel([0.587646, -1.205881, -2.670223, -0.836285, 1.570796, 2.158442],accel_mss,speed_ms,0,blend_radius_m)
  movel([0.584359, -1.207554, -2.669411, -0.835424, 1.570796, 2.155155],accel_mss,speed_ms,0,blend_radius_m)
  movel([0.581016, -1.208886, -2.668762, -0.834741, 1.570796, 2.151812],accel_mss,speed_ms,0,blend_radius_m)
  movel([0.577648, -1.209840, -2.668297, -0.834253, 1.570796, 2.148444],accel_mss,speed_ms,0,blend_radius_m)
  movel([0.575963, -1.209968, -2.668234, -0.834187, 1.570796, 2.146759],accel_mss,speed_ms,0,blend_radius_m)
  movel([0.574295, -1.209824, -2.668304, -0.834261, 1.570796, 2.145091],accel_mss,speed_ms,0,blend_radius_m)
  movel([0.572793, -1.209702, -2.668364, -0.834323, 1.570796, 2.143589],accel_mss,speed_ms,0,blend_radius_m)
  movel([0.571606, -1.209907, -2.668264, -0.834219, 1.570796, 2.142403],accel_mss,speed_ms,0,blend_radius_m)
  movel([0.569556, -1.211331, -2.667566, -0.833492, 1.570796, 2.140352],accel_mss,speed_ms,0,blend_radius_m)
  movel([0.566851, -1.213632, -2.666435, -0.832322, 1.570796, 2.137647],accel_mss,speed_ms,0,blend_radius_m)
  movel([0.564044, -1.216061, -2.665234, -0.831094, 1.570796, 2.134840],accel_mss,speed_ms,0,blend_radius_m)
  movel([0.561677, -1.217879, -2.664330, -0.830179, 1.570796, 2.132473],accel_mss,speed_ms,0,blend_radius_m)
  movel([0.557009, -1.220538, -2.663002, -0.828848, 1.570796, 2.127806],accel_mss,speed_ms,0,blend_radius_m)
  movel([0.552849, -1.222245, -2.662146, -0.827998, 1.570796, 2.123645],accel_mss,speed_ms,0,blend_radius_m)
  movel([0.549147, -1.223088, -2.661722, -0.827579, 1.570796, 2.119944],accel_mss,speed_ms,0,blend_radius_m)
  movel([0.545860, -1.223164, -2.661683, -0.827541, 1.570796, 2.116656],accel_mss,speed_ms,0,blend_radius_m)
  movel([0.542946, -1.222560, -2.661988, -0.827841, 1.570796, 2.113742],accel_mss,speed_ms,0,blend_radius_m)
  movel([0.540365, -1.221359, -2.662591, -0.828439, 1.570796, 2.111161],accel_mss,speed_ms,0,blend_radius_m)
  movel([0.538085, -1.219643, -2.663451, -0.829296, 1.570796, 2.108882],accel_mss,speed_ms,0,blend_radius_m)
  movel([0.536073, -1.217497, -2.664521, -0.830372, 1.570796, 2.106869],accel_mss,speed_ms,0,blend_radius_m)
  movel([0.532697, -1.212253, -2.667114, -0.833022, 1.570796, 2.103494],accel_mss,speed_ms,0,blend_radius_m)
  movel([0.529984, -1.206302, -2.670019, -0.836068, 1.570796, 2.100781],accel_mss,speed_ms,0,blend_radius_m)
  movel([0.525502, -1.195089, -2.675386, -0.841913, 1.570796, 2.096299],accel_mss,speed_ms,0,blend_radius_m)
  movel([0.522928, -1.190586, -2.677503, -0.844300, 1.570796, 2.093724],accel_mss,speed_ms,0,blend_radius_m)
  movel([0.519344, -1.185857, -2.679703, -0.846829, 1.570796, 2.090141],accel_mss,speed_ms,0,blend_radius_m)
  movel([0.514890, -1.181195, -2.681848, -0.849346, 1.570796, 2.085686],accel_mss,speed_ms,0,blend_radius_m)
  movel([0.509718, -1.176896, -2.683805, -0.851688, 1.570796, 2.080514],accel_mss,speed_ms,0,blend_radius_m)
  movel([0.503990, -1.173254, -2.685448, -0.853686, 1.570796, 2.074786],accel_mss,speed_ms,0,blend_radius_m)
  movel([0.497882, -1.170560, -2.686655, -0.855174, 1.570796, 2.068679],accel_mss,speed_ms,0,blend_radius_m)
  movel([0.491590, -1.169090, -2.687310, -0.855989, 1.570796, 2.062387],accel_mss,speed_ms,0,blend_radius_m)
  movel([0.488434, -1.168898, -2.687395, -0.856095, 1.570796, 2.059231],accel_mss,speed_ms,0,blend_radius_m)
  movel([0.485311, -1.169115, -2.687299, -0.855975, 1.570796, 2.056108],accel_mss,speed_ms,0,blend_radius_m)
  movel([0.481950, -1.169764, -2.687010, -0.855615, 1.570796, 2.052746],accel_mss,speed_ms,0,blend_radius_m)
  movel([0.477914, -1.170926, -2.686491, -0.854971, 1.570796, 2.048710],accel_mss,speed_ms,0,blend_radius_m)
  movel([0.473436, -1.172620, -2.685733, -0.854036, 1.570796, 2.044233],accel_mss,speed_ms,0,blend_radius_m)
  movel([0.468754, -1.174864, -2.684724, -0.852801, 1.570796, 2.039551],accel_mss,speed_ms,0,blend_radius_m)
  movel([0.464101, -1.177679, -2.683451, -0.851260, 1.570796, 2.034897],accel_mss,speed_ms,0,blend_radius_m)
  movel([0.459709, -1.181067, -2.681907, -0.849416, 1.570796, 2.030506],accel_mss,speed_ms,0,blend_radius_m)
  movel([0.455816, -1.185032, -2.680084, -0.847273, 1.570796, 2.026613],accel_mss,speed_ms,0,blend_radius_m)
  movel([0.454127, -1.187234, -2.679065, -0.846090, 1.570796, 2.024923],accel_mss,speed_ms,0,blend_radius_m)
  movel([0.452646, -1.189583, -2.677972, -0.844834, 1.570796, 2.023443],accel_mss,speed_ms,0,blend_radius_m)
  movel([0.451023, -1.193247, -2.676255, -0.842887, 1.570796, 2.021820],accel_mss,speed_ms,0,blend_radius_m)
  movel([0.450539, -1.196342, -2.674793, -0.841253, 1.570796, 2.021336],accel_mss,speed_ms,0,blend_radius_m)
  movel([0.451063, -1.198928, -2.673564, -0.839896, 1.570796, 2.021859],accel_mss,speed_ms,0,blend_radius_m)
  movel([0.452469, -1.201057, -2.672547, -0.838785, 1.570796, 2.023265],accel_mss,speed_ms,0,blend_radius_m)
  movel([0.454630, -1.202783, -2.671718, -0.837887, 1.570796, 2.025427],accel_mss,speed_ms,0,blend_radius_m)
  movel([0.457425, -1.204162, -2.671054, -0.837173, 1.570796, 2.028222],accel_mss,speed_ms,0,blend_radius_m)
  movel([0.460733, -1.205240, -2.670533, -0.836616, 1.570796, 2.031529],accel_mss,speed_ms,0,blend_radius_m)
  movel([0.464437, -1.206072, -2.670130, -0.836186, 1.570796, 2.035233],accel_mss,speed_ms,0,blend_radius_m)
  movel([0.472559, -1.207171, -2.669597, -0.835621, 1.570796, 2.043355],accel_mss,speed_ms,0,blend_radius_m)
  movel([0.480857, -1.207811, -2.669286, -0.835292, 1.570796, 2.051654],accel_mss,speed_ms,0,blend_radius_m)
  movel([0.488409, -1.208306, -2.669045, -0.835038, 1.570796, 2.059205],accel_mss,speed_ms,0,blend_radius_m)
  movel([0.494290, -1.208952, -2.668730, -0.834707, 1.570796, 2.065086],accel_mss,speed_ms,0,blend_radius_m)
  movel([0.508074, -1.211290, -2.667586, -0.833512, 1.570796, 2.078870],accel_mss,speed_ms,0,blend_radius_m)
  movel([0.515256, -1.212835, -2.666827, -0.832726, 1.570796, 2.086053],accel_mss,speed_ms,0,blend_radius_m)
  movel([0.520574, -1.214495, -2.666009, -0.831885, 1.570796, 2.091370],accel_mss,speed_ms,0,blend_radius_m)
  movel([0.522393, -1.215497, -2.665513, -0.831379, 1.570796, 2.093189],accel_mss,speed_ms,0,blend_radius_m)
  movel([0.523902, -1.216783, -2.664876, -0.830731, 1.570796, 2.094699],accel_mss,speed_ms,0,blend_radius_m)
  movel([0.526056, -1.220083, -2.663230, -0.829076, 1.570796, 2.096852],accel_mss,speed_ms,0,blend_radius_m)
  movel([0.527136, -1.224176, -2.661173, -0.827040, 1.570796, 2.097932],accel_mss,speed_ms,0,blend_radius_m)
  movel([0.527250, -1.228846, -2.658802, -0.824741, 1.570796, 2.098047],accel_mss,speed_ms,0,blend_radius_m)
  movel([0.526516, -1.233885, -2.656215, -0.822289, 1.570796, 2.097313],accel_mss,speed_ms,0,blend_radius_m)
  movel([0.525036, -1.239090, -2.653512, -0.819786, 1.570796, 2.095833],accel_mss,speed_ms,0,blend_radius_m)
  movel([0.522921, -1.244265, -2.650794, -0.817331, 1.570796, 2.093717],accel_mss,speed_ms,0,blend_radius_m)
  movel([0.520270, -1.249225, -2.648158, -0.815006, 1.570796, 2.091066],accel_mss,speed_ms,0,blend_radius_m)
  movel([0.516302, -1.255024, -2.645039, -0.812326, 1.570796, 2.087098],accel_mss,speed_ms,0,blend_radius_m)
  movel([0.514351, -1.257310, -2.643799, -0.811280, 1.570796, 2.085147],accel_mss,speed_ms,0,blend_radius_m)
  movel([0.512407, -1.259240, -2.642747, -0.810403, 1.570796, 2.083203],accel_mss,speed_ms,0,blend_radius_m)
  movel([0.510454, -1.260861, -2.641859, -0.809669, 1.570796, 2.081250],accel_mss,speed_ms,0,blend_radius_m)
  movel([0.508478, -1.262210, -2.641118, -0.809060, 1.570796, 2.079275],accel_mss,speed_ms,0,blend_radius_m)
  movel([0.504425, -1.264256, -2.639991, -0.808142, 1.570796, 2.075221],accel_mss,speed_ms,0,blend_radius_m)
  movel([0.500148, -1.265695, -2.639194, -0.807500, 1.570796, 2.070944],accel_mss,speed_ms,0,blend_radius_m)
  movel([0.495563, -1.266831, -2.638564, -0.806994, 1.570796, 2.066360],accel_mss,speed_ms,0,blend_radius_m)
  movel([0.485153, -1.269421, -2.637121, -0.805847, 1.570796, 2.055950],accel_mss,speed_ms,0,blend_radius_m)
  movel([0.484610, -1.269606, -2.637017, -0.805766, 1.570796, 2.055407],accel_mss,speed_ms,0,blend_radius_m)
  movel([0.484778, -1.269712, -2.636958, -0.805719, 1.570796, 2.055575],accel_mss,speed_ms,0,blend_radius_m)
  movel([0.486875, -1.269742, -2.636941, -0.805706, 1.570796, 2.057672],accel_mss,speed_ms,0,blend_radius_m)
  movel([0.495499, -1.269356, -2.637157, -0.805876, 1.570796, 2.066296],accel_mss,speed_ms,0,blend_radius_m)
  movel([0.509774, -1.268838, -2.637446, -0.806105, 1.570796, 2.080571],accel_mss,speed_ms,0,blend_radius_m)
  movel([0.501277, -1.272786, -2.635233, -0.804370, 1.570796, 2.072074],accel_mss,speed_ms,0,blend_radius_m)
  movel([0.491841, -1.276761, -2.632985, -0.802642, 1.570796, 2.062638],accel_mss,speed_ms,0,blend_radius_m)
  movel([0.481807, -1.280688, -2.630746, -0.800955, 1.570796, 2.052604],accel_mss,speed_ms,0,blend_radius_m)
  movel([0.471511, -1.284482, -2.628563, -0.799343, 1.570796, 2.042307],accel_mss,speed_ms,0,blend_radius_m)
  movel([0.451457, -1.291297, -2.624598, -0.796494, 1.570796, 2.022254],accel_mss,speed_ms,0,blend_radius_m)
  movel([0.442351, -1.294110, -2.622943, -0.795335, 1.570796, 2.013147],accel_mss,speed_ms,0,blend_radius_m)
  movel([0.434287, -1.296377, -2.621603, -0.794409, 1.570796, 2.005083],accel_mss,speed_ms,0,blend_radius_m)
  movel([0.422943, -1.303775, -2.617182, -0.791431, 1.570796, 1.993739],accel_mss,speed_ms,0,blend_radius_m)
  movel([0.411504, -1.311826, -2.612291, -0.788272, 1.570796, 1.982300],accel_mss,speed_ms,0,blend_radius_m)
  movel([0.388708, -1.328733, -2.601742, -0.781914, 1.570796, 1.959504],accel_mss,speed_ms,0,blend_radius_m)
  movel([0.377505, -1.337050, -2.596412, -0.778927, 1.570796, 1.948301],accel_mss,speed_ms,0,blend_radius_m)
  movel([0.366504, -1.344945, -2.591265, -0.776178, 1.570796, 1.937301],accel_mss,speed_ms,0,blend_radius_m)
  movel([0.355748, -1.352184, -2.586471, -0.773733, 1.570796, 1.926544],accel_mss,speed_ms,0,blend_radius_m)
  movel([0.345262, -1.358551, -2.582195, -0.771643, 1.570796, 1.916058],accel_mss,speed_ms,0,blend_radius_m)
  movel([0.341198, -1.360699, -2.580740, -0.770950, 1.570796, 1.911994],accel_mss,speed_ms,0,blend_radius_m)
  movel([0.337339, -1.362432, -2.579561, -0.770396, 1.570796, 1.908136],accel_mss,speed_ms,0,blend_radius_m)
  movel([0.333707, -1.363755, -2.578658, -0.769976, 1.570796, 1.904503],accel_mss,speed_ms,0,blend_radius_m)
  movel([0.330321, -1.364673, -2.578030, -0.769686, 1.570796, 1.901117],accel_mss,speed_ms,0,blend_radius_m)
  movel([0.327200, -1.365186, -2.577678, -0.769525, 1.570796, 1.897996],accel_mss,speed_ms,0,blend_radius_m)
  movel([0.324365, -1.365298, -2.577602, -0.769489, 1.570796, 1.895161],accel_mss,speed_ms,0,blend_radius_m)
  movel([0.321836, -1.365008, -2.577801, -0.769581, 1.570796, 1.892632],accel_mss,speed_ms,0,blend_radius_m)
  movel([0.319635, -1.364317, -2.578274, -0.769799, 1.570796, 1.890432],accel_mss,speed_ms,0,blend_radius_m)
  movel([0.317785, -1.363222, -2.579021, -0.770145, 1.570796, 1.888582],accel_mss,speed_ms,0,blend_radius_m)
  movel([0.316314, -1.361721, -2.580045, -0.770623, 1.570796, 1.887110],accel_mss,speed_ms,0,blend_radius_m)
  movel([0.315242, -1.359812, -2.581341, -0.771236, 1.570796, 1.886038],accel_mss,speed_ms,0,blend_radius_m)
  movel([0.314595, -1.357494, -2.582909, -0.771986, 1.570796, 1.885391],accel_mss,speed_ms,0,blend_radius_m)
  movel([0.314408, -1.354754, -2.584752, -0.772883, 1.570796, 1.885204],accel_mss,speed_ms,0,blend_radius_m)
  movel([0.314703, -1.351593, -2.586865, -0.773930, 1.570796, 1.885499],accel_mss,speed_ms,0,blend_radius_m)
  movel([0.315513, -1.348002, -2.589250, -0.775137, 1.570796, 1.886310],accel_mss,speed_ms,0,blend_radius_m)
  movel([0.316873, -1.343972, -2.591904, -0.776513, 1.570796, 1.887669],accel_mss,speed_ms,0,blend_radius_m)
  movel([0.320026, -1.345111, -2.591156, -0.776122, 1.570796, 1.890822],accel_mss,speed_ms,0,blend_radius_m)
  movel([0.321631, -1.345562, -2.590860, -0.775968, 1.570796, 1.892428],accel_mss,speed_ms,0,blend_radius_m)
  movel([0.323409, -1.345574, -2.590852, -0.775963, 1.570796, 1.894205],accel_mss,speed_ms,0,blend_radius_m)
  movel([0.324957, -1.345102, -2.591162, -0.776125, 1.570796, 1.895753],accel_mss,speed_ms,0,blend_radius_m)
  movel([0.326886, -1.344144, -2.591791, -0.776454, 1.570796, 1.897682],accel_mss,speed_ms,0,blend_radius_m)
  movel([0.331685, -1.341013, -2.593839, -0.777537, 1.570796, 1.902482],accel_mss,speed_ms,0,blend_radius_m)
  movel([0.337409, -1.336650, -2.596670, -0.779068, 1.570796, 1.908205],accel_mss,speed_ms,0,blend_radius_m)
  movel([0.343643, -1.331525, -2.599963, -0.780901, 1.570796, 1.914439],accel_mss,speed_ms,0,blend_radius_m)
  movel([0.355929, -1.320912, -2.606669, -0.784808, 1.570796, 1.926725],accel_mss,speed_ms,0,blend_radius_m)
  movel([0.364909, -1.313157, -2.611475, -0.787757, 1.570796, 1.935705],accel_mss,speed_ms,0,blend_radius_m)
  movel([0.372993, -1.306914, -2.615285, -0.790189, 1.570796, 1.943789],accel_mss,speed_ms,0,blend_radius_m)
  movel([0.381163, -1.300641, -2.619064, -0.792684, 1.570796, 1.951960],accel_mss,speed_ms,0,blend_radius_m)
  movel([0.364737, -1.304066, -2.617008, -0.791316, 1.570796, 1.935533],accel_mss,speed_ms,0,blend_radius_m)
  movel([0.356262, -1.305520, -2.616130, -0.790739, 1.570796, 1.927058],accel_mss,speed_ms,0,blend_radius_m)
  movel([0.348215, -1.306218, -2.615707, -0.790463, 1.570796, 1.919012],accel_mss,speed_ms,0,blend_radius_m)
  movel([0.344490, -1.306142, -2.615754, -0.790494, 1.570796, 1.915286],accel_mss,speed_ms,0,blend_radius_m)
  movel([0.341037, -1.305708, -2.616016, -0.790665, 1.570796, 1.911833],accel_mss,speed_ms,0,blend_radius_m)
  movel([0.337907, -1.304857, -2.616530, -0.791002, 1.570796, 1.908703],accel_mss,speed_ms,0,blend_radius_m)
  movel([0.335155, -1.303530, -2.617330, -0.791529, 1.570796, 1.905951],accel_mss,speed_ms,0,blend_radius_m)
  movel([0.332839, -1.301665, -2.618450, -0.792273, 1.570796, 1.903635],accel_mss,speed_ms,0,blend_radius_m)
  movel([0.331018, -1.299196, -2.619927, -0.793266, 1.570796, 1.901814],accel_mss,speed_ms,0,blend_radius_m)
  movel([0.329744, -1.296061, -2.621791, -0.794538, 1.570796, 1.900540],accel_mss,speed_ms,0,blend_radius_m)
  movel([0.329083, -1.292183, -2.624078, -0.796128, 1.570796, 1.899879],accel_mss,speed_ms,0,blend_radius_m)
  movel([0.329274, -1.287156, -2.627015, -0.798219, 1.570796, 1.900071],accel_mss,speed_ms,0,blend_radius_m)
  movel([0.330527, -1.281649, -2.630195, -0.800545, 1.570796, 1.901324],accel_mss,speed_ms,0,blend_radius_m)
  movel([0.332760, -1.275831, -2.633513, -0.803045, 1.570796, 1.903556],accel_mss,speed_ms,0,blend_radius_m)
  movel([0.335886, -1.269885, -2.636861, -0.805643, 1.570796, 1.906682],accel_mss,speed_ms,0,blend_radius_m)
  movel([0.339813, -1.264003, -2.640130, -0.808256, 1.570796, 1.910609],accel_mss,speed_ms,0,blend_radius_m)
  movel([0.344441, -1.258385, -2.643213, -0.810791, 1.570796, 1.915237],accel_mss,speed_ms,0,blend_radius_m)
  movel([0.349662, -1.253238, -2.646004, -0.813147, 1.570796, 1.920459],accel_mss,speed_ms,0,blend_radius_m)
  movel([0.355368, -1.248780, -2.648395, -0.815213, 1.570796, 1.926164],accel_mss,speed_ms,0,blend_radius_m)
  movel([0.358633, -1.247037, -2.649324, -0.816028, 1.570796, 1.929430],accel_mss,speed_ms,0,blend_radius_m)
  movel([0.362267, -1.245798, -2.649982, -0.816609, 1.570796, 1.933064],accel_mss,speed_ms,0,blend_radius_m)
  movel([0.365103, -1.245534, -2.650122, -0.816733, 1.570796, 1.935899],accel_mss,speed_ms,0,blend_radius_m)
  movel([0.365856, -1.245904, -2.649926, -0.816559, 1.570796, 1.936653],accel_mss,speed_ms,0,blend_radius_m)
  movel([0.365974, -1.246687, -2.649510, -0.816192, 1.570796, 1.936770],accel_mss,speed_ms,0,blend_radius_m)
  movel([0.363106, -1.247613, -2.649018, -0.815758, 1.570796, 1.933903],accel_mss,speed_ms,0,blend_radius_m)
  movel([0.360648, -1.248698, -2.648439, -0.815252, 1.570796, 1.931444],accel_mss,speed_ms,0,blend_radius_m)
  movel([0.358588, -1.249914, -2.647790, -0.814686, 1.570796, 1.929384],accel_mss,speed_ms,0,blend_radius_m)
  movel([0.356915, -1.251229, -2.647085, -0.814075, 1.570796, 1.927711],accel_mss,speed_ms,0,blend_radius_m)
  movel([0.355611, -1.252620, -2.646337, -0.813432, 1.570796, 1.926408],accel_mss,speed_ms,0,blend_radius_m)
  movel([0.354669, -1.254059, -2.645561, -0.812769, 1.570796, 1.925465],accel_mss,speed_ms,0,blend_radius_m)
  movel([0.354068, -1.255517, -2.644772, -0.812100, 1.570796, 1.924865],accel_mss,speed_ms,0,blend_radius_m)
  movel([0.353797, -1.256972, -2.643982, -0.811434, 1.570796, 1.924593],accel_mss,speed_ms,0,blend_radius_m)
  movel([0.354183, -1.259776, -2.642454, -0.810160, 1.570796, 1.924979],accel_mss,speed_ms,0,blend_radius_m)
  movel([0.355701, -1.262277, -2.641082, -0.809031, 1.570796, 1.926497],accel_mss,speed_ms,0,blend_radius_m)
  movel([0.358242, -1.264286, -2.639974, -0.808129, 1.570796, 1.929038],accel_mss,speed_ms,0,blend_radius_m)
  movel([0.361695, -1.265617, -2.639237, -0.807534, 1.570796, 1.932492],accel_mss,speed_ms,0,blend_radius_m)
  movel([0.364100, -1.265932, -2.639063, -0.807394, 1.570796, 1.934896],accel_mss,speed_ms,0,blend_radius_m)
  movel([0.367189, -1.265929, -2.639065, -0.807396, 1.570796, 1.937985],accel_mss,speed_ms,0,blend_radius_m)
  movel([0.375053, -1.265116, -2.639515, -0.807758, 1.570796, 1.945849],accel_mss,speed_ms,0,blend_radius_m)
  movel([0.384568, -1.263485, -2.640416, -0.808488, 1.570796, 1.955364],accel_mss,speed_ms,0,blend_radius_m)
  movel([0.395013, -1.261330, -2.641602, -0.809457, 1.570796, 1.965809],accel_mss,speed_ms,0,blend_radius_m)
  movel([0.415806, -1.256499, -2.644240, -0.811651, 1.570796, 1.986602],accel_mss,speed_ms,0,blend_radius_m)
  movel([0.431593, -1.252551, -2.646374, -0.813464, 1.570796, 2.002390],accel_mss,speed_ms,0,blend_radius_m)
  movel([0.439550, -1.250558, -2.647445, -0.814386, 1.570796, 2.010346],accel_mss,speed_ms,0,blend_radius_m)
  movel([0.443868, -1.249342, -2.648096, -0.814952, 1.570796, 2.014664],accel_mss,speed_ms,0,blend_radius_m)
  movel([0.447186, -1.248121, -2.648747, -0.815521, 1.570796, 2.017982],accel_mss,speed_ms,0,blend_radius_m)
  movel([0.448107, -1.247593, -2.649028, -0.815768, 1.570796, 2.018903],accel_mss,speed_ms,0,blend_radius_m)
  movel([0.448491, -1.247123, -2.649278, -0.815987, 1.570796, 2.019287],accel_mss,speed_ms,0,blend_radius_m)
  movel([0.448096, -1.246077, -2.649834, -0.816478, 1.570796, 2.018893],accel_mss,speed_ms,0,blend_radius_m)
  movel([0.445706, -1.243973, -2.650948, -0.817468, 1.570796, 2.016503],accel_mss,speed_ms,0,blend_radius_m)
  movel([0.442615, -1.242449, -2.651751, -0.818189, 1.570796, 2.013412],accel_mss,speed_ms,0,blend_radius_m)
  movel([0.435646, -1.239588, -2.653252, -0.819549, 1.570796, 2.006443],accel_mss,speed_ms,0,blend_radius_m)
  movel([0.432418, -1.237456, -2.654364, -0.820569, 1.570796, 2.003214],accel_mss,speed_ms,0,blend_radius_m)
  movel([0.429795, -1.234313, -2.655994, -0.822082, 1.570796, 2.000591],accel_mss,speed_ms,0,blend_radius_m)
  movel([0.428813, -1.232228, -2.657069, -0.823092, 1.570796, 1.999610],accel_mss,speed_ms,0,blend_radius_m)
  movel([0.428108, -1.229731, -2.658350, -0.824308, 1.570796, 1.998904],accel_mss,speed_ms,0,blend_radius_m)
  movel([0.427720, -1.226759, -2.659864, -0.825765, 1.570796, 1.998516],accel_mss,speed_ms,0,blend_radius_m)
  movel([0.427696, -1.223259, -2.661635, -0.827494, 1.570796, 1.998493],accel_mss,speed_ms,0,blend_radius_m)
  movel([0.428383, -1.218343, -2.664099, -0.829947, 1.570796, 1.999179],accel_mss,speed_ms,0,blend_radius_m)
  movel([0.429937, -1.213396, -2.666551, -0.832442, 1.570796, 2.000733],accel_mss,speed_ms,0,blend_radius_m)
  movel([0.432257, -1.208442, -2.668979, -0.834968, 1.570796, 2.003053],accel_mss,speed_ms,0,blend_radius_m)
  movel([0.435250, -1.203501, -2.671373, -0.837515, 1.570796, 2.006046],accel_mss,speed_ms,0,blend_radius_m)
  movel([0.438815, -1.198593, -2.673724, -0.840072, 1.570796, 2.009611],accel_mss,speed_ms,0,blend_radius_m)
  movel([0.442846, -1.193743, -2.676021, -0.842624, 1.570796, 2.013642],accel_mss,speed_ms,0,blend_radius_m)
  movel([0.447238, -1.188978, -2.678254, -0.845157, 1.570796, 2.018034],accel_mss,speed_ms,0,blend_radius_m)
  movel([0.451880, -1.184320, -2.680413, -0.847656, 1.570796, 2.022676],accel_mss,speed_ms,0,blend_radius_m)
  movel([0.461042, -1.176089, -2.684170, -0.852129, 1.570796, 2.031839],accel_mss,speed_ms,0,blend_radius_m)
  movel([0.469454, -1.169622, -2.687073, -0.855694, 1.570796, 2.040250],accel_mss,speed_ms,0,blend_radius_m)
  movel([0.476694, -1.164844, -2.689190, -0.858355, 1.570796, 2.047490],accel_mss,speed_ms,0,blend_radius_m)
  movel([0.482357, -1.161662, -2.690586, -0.860141, 1.570796, 2.053153],accel_mss,speed_ms,0,blend_radius_m)
  movel([0.490737, -1.157933, -2.692209, -0.862246, 1.570796, 2.061533],accel_mss,speed_ms,0,blend_radius_m)
  movel([0.498778, -1.155444, -2.693285, -0.863660, 1.570796, 2.069574],accel_mss,speed_ms,0,blend_radius_m)
  movel([0.506373, -1.154176, -2.693831, -0.864383, 1.570796, 2.077169],accel_mss,speed_ms,0,blend_radius_m)
  movel([0.513424, -1.154101, -2.693863, -0.864425, 1.570796, 2.084220],accel_mss,speed_ms,0,blend_radius_m)
  movel([0.519834, -1.155174, -2.693401, -0.863814, 1.570796, 2.090631],accel_mss,speed_ms,0,blend_radius_m)
  movel([0.525516, -1.157346, -2.692464, -0.862579, 1.570796, 2.096312],accel_mss,speed_ms,0,blend_radius_m)
  movel([0.530388, -1.160561, -2.691067, -0.860761, 1.570796, 2.101184],accel_mss,speed_ms,0,blend_radius_m)
  movel([0.534374, -1.164753, -2.689230, -0.858406, 1.570796, 2.105170],accel_mss,speed_ms,0,blend_radius_m)
  movel([0.537149, -1.169301, -2.687216, -0.855872, 1.570796, 2.107945],accel_mss,speed_ms,0,blend_radius_m)
  movel([0.539381, -1.174243, -2.685003, -0.853142, 1.570796, 2.110177],accel_mss,speed_ms,0,blend_radius_m)
  movel([0.541475, -1.179168, -2.682773, -0.850448, 1.570796, 2.112272],accel_mss,speed_ms,0,blend_radius_m)
  movel([0.543831, -1.183677, -2.680709, -0.848003, 1.570796, 2.114627],accel_mss,speed_ms,0,blend_radius_m)
  movel([0.546842, -1.187393, -2.678991, -0.846005, 1.570796, 2.117638],accel_mss,speed_ms,0,blend_radius_m)
  movel([0.548716, -1.188833, -2.678322, -0.845234, 1.570796, 2.119513],accel_mss,speed_ms,0,blend_radius_m)
  movel([0.550899, -1.189937, -2.677807, -0.844645, 1.570796, 2.121695],accel_mss,speed_ms,0,blend_radius_m)
  movel([0.553441, -1.190662, -2.677468, -0.844259, 1.570796, 2.124238],accel_mss,speed_ms,0,blend_radius_m)
  movel([0.556397, -1.190954, -2.677331, -0.844103, 1.570796, 2.127194],accel_mss,speed_ms,0,blend_radius_m)
  movel([0.559817, -1.190777, -2.677414, -0.844198, 1.570796, 2.130613],accel_mss,speed_ms,0,blend_radius_m)
  movel([0.563749, -1.190080, -2.677740, -0.844569, 1.570796, 2.134545],accel_mss,speed_ms,0,blend_radius_m)
  movel([0.567343, -1.188924, -2.678279, -0.845186, 1.570796, 2.138139],accel_mss,speed_ms,0,blend_radius_m)
  movel([0.570516, -1.187275, -2.679046, -0.846068, 1.570796, 2.141313],accel_mss,speed_ms,0,blend_radius_m)
  movel([0.573266, -1.185225, -2.679995, -0.847169, 1.570796, 2.144063],accel_mss,speed_ms,0,blend_radius_m)
  movel([0.575583, -1.182870, -2.681080, -0.848439, 1.570796, 2.146379],accel_mss,speed_ms,0,blend_radius_m)
  movel([0.577458, -1.180310, -2.682252, -0.849826, 1.570796, 2.148255],accel_mss,speed_ms,0,blend_radius_m)
  movel([0.578887, -1.177643, -2.683467, -0.851279, 1.570796, 2.149683],accel_mss,speed_ms,0,blend_radius_m)
  movel([0.579854, -1.174973, -2.684675, -0.852741, 1.570796, 2.150650],accel_mss,speed_ms,0,blend_radius_m)
  movel([0.580343, -1.172405, -2.685829, -0.854154, 1.570796, 2.151140],accel_mss,speed_ms,0,blend_radius_m)
  movel([0.580340, -1.170051, -2.686882, -0.855456, 1.570796, 2.151137],accel_mss,speed_ms,0,blend_radius_m)
  movel([0.579838, -1.168016, -2.687787, -0.856586, 1.570796, 2.150634],accel_mss,speed_ms,0,blend_radius_m)
  movel([0.578818, -1.166414, -2.688497, -0.857478, 1.570796, 2.149615],accel_mss,speed_ms,0,blend_radius_m)
  movel([0.577270, -1.165356, -2.688964, -0.858069, 1.570796, 2.148067],accel_mss,speed_ms,0,blend_radius_m)
  movel([0.575187, -1.164951, -2.689143, -0.858295, 1.570796, 2.145983],accel_mss,speed_ms,0,blend_radius_m)
  movel([0.572561, -1.165309, -2.688985, -0.858095, 1.570796, 2.143357],accel_mss,speed_ms,0,blend_radius_m)
  movel([0.569385, -1.166537, -2.688443, -0.857410, 1.570796, 2.140181],accel_mss,speed_ms,0,blend_radius_m)
  movel([0.565666, -1.168733, -2.687469, -0.856187, 1.570796, 2.136462],accel_mss,speed_ms,0,blend_radius_m)
  movel([0.567625, -1.169139, -2.687288, -0.855962, 1.570796, 2.138421],accel_mss,speed_ms,0,blend_radius_m)
  movel([0.568986, -1.169951, -2.686926, -0.855511, 1.570796, 2.139782],accel_mss,speed_ms,0,blend_radius_m)
  movel([0.569746, -1.171108, -2.686410, -0.854871, 1.570796, 2.140543],accel_mss,speed_ms,0,blend_radius_m)
  movel([0.569899, -1.172542, -2.685768, -0.854079, 1.570796, 2.140696],accel_mss,speed_ms,0,blend_radius_m)
  movel([0.569435, -1.174199, -2.685024, -0.853166, 1.570796, 2.140232],accel_mss,speed_ms,0,blend_radius_m)
  movel([0.568358, -1.176014, -2.684205, -0.852170, 1.570796, 2.139154],accel_mss,speed_ms,0,blend_radius_m)
  movel([0.566658, -1.177932, -2.683335, -0.851121, 1.570796, 2.137455],accel_mss,speed_ms,0,blend_radius_m)
  movel([0.564334, -1.179892, -2.682443, -0.850054, 1.570796, 2.135130],accel_mss,speed_ms,0,blend_radius_m)
  movel([0.560104, -1.182534, -2.681234, -0.848621, 1.570796, 2.130901],accel_mss,speed_ms,0,blend_radius_m)
  movel([0.556297, -1.183951, -2.680583, -0.847855, 1.570796, 2.127094],accel_mss,speed_ms,0,blend_radius_m)
  movel([0.552930, -1.184268, -2.680437, -0.847684, 1.570796, 2.123727],accel_mss,speed_ms,0,blend_radius_m)
  movel([0.550026, -1.183600, -2.680744, -0.848045, 1.570796, 2.120822],accel_mss,speed_ms,0,blend_radius_m)
  movel([0.547608, -1.182068, -2.681448, -0.848873, 1.570796, 2.118404],accel_mss,speed_ms,0,blend_radius_m)
  movel([0.545712, -1.179770, -2.682499, -0.850120, 1.570796, 2.116508],accel_mss,speed_ms,0,blend_radius_m)
  movel([0.544366, -1.176817, -2.683841, -0.851731, 1.570796, 2.115163],accel_mss,speed_ms,0,blend_radius_m)
  movel([0.543618, -1.173310, -2.685424, -0.853656, 1.570796, 2.114414],accel_mss,speed_ms,0,blend_radius_m)
  movel([0.543498, -1.169355, -2.687192, -0.855842, 1.570796, 2.114295],accel_mss,speed_ms,0,blend_radius_m)
  movel([0.544057, -1.165059, -2.689095, -0.858235, 1.570796, 2.114854],accel_mss,speed_ms,0,blend_radius_m)
  movel([0.545334, -1.160528, -2.691081, -0.860780, 1.570796, 2.116131],accel_mss,speed_ms,0,blend_radius_m)
  movel([0.547380, -1.155871, -2.693101, -0.863417, 1.570796, 2.118176],accel_mss,speed_ms,0,blend_radius_m)
  movel([0.550233, -1.151211, -2.695100, -0.866078, 1.570796, 2.121029],accel_mss,speed_ms,0,blend_radius_m)
  movel([0.553938, -1.146667, -2.697028, -0.868694, 1.570796, 2.124735],accel_mss,speed_ms,0,blend_radius_m)
  movel([0.558537, -1.142369, -2.698833, -0.871187, 1.570796, 2.129333],accel_mss,speed_ms,0,blend_radius_m)
  movel([0.564060, -1.138457, -2.700460, -0.873472, 1.570796, 2.134857],accel_mss,speed_ms,0,blend_radius_m)
  movel([0.568167, -1.136126, -2.701422, -0.874841, 1.570796, 2.138963],accel_mss,speed_ms,0,blend_radius_m)
  movel([0.572245, -1.134166, -2.702227, -0.875996, 1.570796, 2.143042],accel_mss,speed_ms,0,blend_radius_m)
  movel([0.576258, -1.132594, -2.702870, -0.876925, 1.570796, 2.147054],accel_mss,speed_ms,0,blend_radius_m)
  movel([0.580176, -1.131411, -2.703352, -0.877626, 1.570796, 2.150972],accel_mss,speed_ms,0,blend_radius_m)
  movel([0.583954, -1.130630, -2.703670, -0.878090, 1.570796, 2.154750],accel_mss,speed_ms,0,blend_radius_m)
  movel([0.587564, -1.130252, -2.703823, -0.878314, 1.570796, 2.158361],accel_mss,speed_ms,0,blend_radius_m)
  movel([0.590968, -1.130286, -2.703809, -0.878294, 1.570796, 2.161764],accel_mss,speed_ms,0,blend_radius_m)
  movel([0.594134, -1.130733, -2.703628, -0.878028, 1.570796, 2.164930],accel_mss,speed_ms,0,blend_radius_m)
  movel([0.597028, -1.131597, -2.703276, -0.877515, 1.570796, 2.167824],accel_mss,speed_ms,0,blend_radius_m)
  movel([0.599616, -1.132876, -2.702755, -0.876758, 1.570796, 2.170412],accel_mss,speed_ms,0,blend_radius_m)
  movel([0.601866, -1.134574, -2.702060, -0.875755, 1.570796, 2.172663],accel_mss,speed_ms,0,blend_radius_m)
  movel([0.603755, -1.136683, -2.701193, -0.874514, 1.570796, 2.174552],accel_mss,speed_ms,0,blend_radius_m)
  movel([0.605248, -1.139204, -2.700150, -0.873034, 1.570796, 2.176044],accel_mss,speed_ms,0,blend_radius_m)
  movel([0.606317, -1.142132, -2.698932, -0.871325, 1.570796, 2.177114],accel_mss,speed_ms,0,blend_radius_m)
  movel([0.606937, -1.145466, -2.697534, -0.869389, 1.570796, 2.177733],accel_mss,speed_ms,0,blend_radius_m)
  movel([0.607087, -1.149190, -2.695960, -0.867239, 1.570796, 2.177883],accel_mss,speed_ms,0,blend_radius_m)
  movel([0.606291, -1.153310, -2.694202, -0.864877, 1.570796, 2.177088],accel_mss,speed_ms,0,blend_radius_m)
  movel([0.604664, -1.157998, -2.692182, -0.862210, 1.570796, 2.175460],accel_mss,speed_ms,0,blend_radius_m)
  movel([0.603065, -1.162062, -2.690411, -0.859916, 1.570796, 2.173862],accel_mss,speed_ms,0,blend_radius_m)
  movel([0.602340, -1.164334, -2.689414, -0.858641, 1.570796, 2.173136],accel_mss,speed_ms,0,blend_radius_m)
  movel([0.603117, -1.165463, -2.688917, -0.858009, 1.570796, 2.173914],accel_mss,speed_ms,0,blend_radius_m)
  movel([0.604906, -1.166808, -2.688323, -0.857259, 1.570796, 2.175702],accel_mss,speed_ms,0,blend_radius_m)
  movel([0.606874, -1.168291, -2.687665, -0.856433, 1.570796, 2.177671],accel_mss,speed_ms,0,blend_radius_m)
  movel([0.608206, -1.169820, -2.686985, -0.855584, 1.570796, 2.179003],accel_mss,speed_ms,0,blend_radius_m)
  movel([0.609148, -1.172499, -2.685787, -0.854103, 1.570796, 2.179944],accel_mss,speed_ms,0,blend_radius_m)
  movel([0.609507, -1.175355, -2.684502, -0.852532, 1.570796, 2.180304],accel_mss,speed_ms,0,blend_radius_m)
  movel([0.609332, -1.178339, -2.683151, -0.850899, 1.570796, 2.180128],accel_mss,speed_ms,0,blend_radius_m)
  movel([0.608669, -1.181406, -2.681751, -0.849232, 1.570796, 2.179465],accel_mss,speed_ms,0,blend_radius_m)
  movel([0.607559, -1.184511, -2.680325, -0.847554, 1.570796, 2.178356],accel_mss,speed_ms,0,blend_radius_m)
  movel([0.606047, -1.187610, -2.678890, -0.845888, 1.570796, 2.176843],accel_mss,speed_ms,0,blend_radius_m)
  movel([0.604177, -1.190664, -2.677467, -0.844258, 1.570796, 2.174973],accel_mss,speed_ms,0,blend_radius_m)
  movel([0.601988, -1.193635, -2.676073, -0.842682, 1.570796, 2.172784],accel_mss,speed_ms,0,blend_radius_m)
  movel([0.599520, -1.196480, -2.674728, -0.841181, 1.570796, 2.170316],accel_mss,speed_ms,0,blend_radius_m)
  movel([0.596813, -1.199165, -2.673451, -0.839772, 1.570796, 2.167609],accel_mss,speed_ms,0,blend_radius_m)
  movel([0.593907, -1.201650, -2.672262, -0.838476, 1.570796, 2.164704],accel_mss,speed_ms,0,blend_radius_m)
  speed_ms = 0.003
  movel([0.593907, -1.194457, -2.668646, -0.849286, 1.570796, 2.164704],accel_mss,speed_ms,0,blend_radius_m)
  speed_ms = 0.01
  movel([0.593907, -1.167128, -2.653928, -0.891333, 1.570796, 2.164704],accel_mss,speed_ms,0,blend_radius_m)
  #M_RunCode9
  movel([0.613006, -1.166119, -2.654391, -0.891880, 1.570796, 2.183802],accel_mss,speed_ms,0,blend_radius_m)
  #M_RunCode3
  movel([0.613006, -1.193454, -2.669122, -0.849813, 1.570796, 2.183802],accel_mss,speed_ms,0,blend_radius_m)
  speed_ms = 0.003
  movel([0.613006, -1.200650, -2.672742, -0.838997, 1.570796, 2.183802],accel_mss,speed_ms,0,blend_radius_m)
  speed_ms = 0.007
  movel([0.614231, -1.198073, -2.673972, -0.840345, 1.570796, 2.185027],accel_mss,speed_ms,0,blend_radius_m)
  movel([0.617381, -1.192832, -2.676450, -0.843107, 1.570796, 2.188177],accel_mss,speed_ms,0,blend_radius_m)
  movel([0.620239, -1.187690, -2.678853, -0.845846, 1.570796, 2.191036],accel_mss,speed_ms,0,blend_radius_m)
  movel([0.621098, -1.185233, -2.679991, -0.847164, 1.570796, 2.191894],accel_mss,speed_ms,0,blend_radius_m)
  movel([0.621319, -1.182901, -2.681066, -0.848422, 1.570796, 2.192115],accel_mss,speed_ms,0,blend_radius_m)
  movel([0.621745, -1.184314, -2.680416, -0.847660, 1.570796, 2.192541],accel_mss,speed_ms,0,blend_radius_m)
  movel([0.621878, -1.187217, -2.679073, -0.846099, 1.570796, 2.192674],accel_mss,speed_ms,0,blend_radius_m)
  movel([0.621252, -1.190174, -2.677696, -0.844519, 1.570796, 2.192048],accel_mss,speed_ms,0,blend_radius_m)
  movel([0.620104, -1.193169, -2.676292, -0.842928, 1.570796, 2.190901],accel_mss,speed_ms,0,blend_radius_m)
  movel([0.618668, -1.196184, -2.674868, -0.841336, 1.570796, 2.189464],accel_mss,speed_ms,0,blend_radius_m)
  movel([0.615868, -1.202220, -2.671989, -0.838180, 1.570796, 2.186664],accel_mss,speed_ms,0,blend_radius_m)
  movel([0.614962, -1.205209, -2.670548, -0.836632, 1.570796, 2.185759],accel_mss,speed_ms,0,blend_radius_m)
  movel([0.614686, -1.208163, -2.669115, -0.835111, 1.570796, 2.185482],accel_mss,speed_ms,0,blend_radius_m)
  movel([0.615072, -1.211190, -2.667635, -0.833563, 1.570796, 2.185868],accel_mss,speed_ms,0,blend_radius_m)
  movel([0.615450, -1.212711, -2.666888, -0.832789, 1.570796, 2.186246],accel_mss,speed_ms,0,blend_radius_m)
  movel([0.615915, -1.213433, -2.666533, -0.832423, 1.570796, 2.186711],accel_mss,speed_ms,0,blend_radius_m)
  movel([0.617595, -1.212840, -2.666825, -0.832724, 1.570796, 2.188391],accel_mss,speed_ms,0,blend_radius_m)
  movel([0.618968, -1.212419, -2.667032, -0.832938, 1.570796, 2.189764],accel_mss,speed_ms,0,blend_radius_m)
  movel([0.620305, -1.212269, -2.667106, -0.833014, 1.570796, 2.191101],accel_mss,speed_ms,0,blend_radius_m)
  movel([0.622669, -1.212621, -2.666932, -0.832835, 1.570796, 2.193465],accel_mss,speed_ms,0,blend_radius_m)
  movel([0.624193, -1.213319, -2.666589, -0.832481, 1.570796, 2.194990],accel_mss,speed_ms,0,blend_radius_m)
  movel([0.625062, -1.214317, -2.666097, -0.831975, 1.570796, 2.195858],accel_mss,speed_ms,0,blend_radius_m)
  movel([0.625449, -1.215574, -2.665475, -0.831340, 1.570796, 2.196245],accel_mss,speed_ms,0,blend_radius_m)
  movel([0.625510, -1.218680, -2.663931, -0.829778, 1.570796, 2.196306],accel_mss,speed_ms,0,blend_radius_m)
  movel([0.625791, -1.222303, -2.662117, -0.827969, 1.570796, 2.196587],accel_mss,speed_ms,0,blend_radius_m)
  movel([0.627077, -1.226675, -2.659907, -0.825807, 1.570796, 2.197873],accel_mss,speed_ms,0,blend_radius_m)
  movel([0.628549, -1.230884, -2.657759, -0.823746, 1.570796, 2.199345],accel_mss,speed_ms,0,blend_radius_m)
  movel([0.629761, -1.235223, -2.655523, -0.821642, 1.570796, 2.200558],accel_mss,speed_ms,0,blend_radius_m)
  movel([0.630272, -1.239969, -2.653053, -0.819367, 1.570796, 2.201068],accel_mss,speed_ms,0,blend_radius_m)
  movel([0.630087, -1.242744, -2.651596, -0.818049, 1.570796, 2.200883],accel_mss,speed_ms,0,blend_radius_m)
  movel([0.629571, -1.245612, -2.650081, -0.816696, 1.570796, 2.200367],accel_mss,speed_ms,0,blend_radius_m)
  movel([0.627894, -1.251491, -2.646944, -0.813954, 1.570796, 2.198690],accel_mss,speed_ms,0,blend_radius_m)
  movel([0.625907, -1.257332, -2.643787, -0.811270, 1.570796, 2.196704],accel_mss,speed_ms,0,blend_radius_m)
  movel([0.624263, -1.262871, -2.640755, -0.808764, 1.570796, 2.195059],accel_mss,speed_ms,0,blend_radius_m)
  movel([0.622675, -1.271702, -2.635843, -0.804844, 1.570796, 2.193471],accel_mss,speed_ms,0,blend_radius_m)
  movel([0.622103, -1.275427, -2.633742, -0.803220, 1.570796, 2.192899],accel_mss,speed_ms,0,blend_radius_m)
  movel([0.621328, -1.278990, -2.631717, -0.801683, 1.570796, 2.192124],accel_mss,speed_ms,0,blend_radius_m)
  movel([0.620089, -1.282605, -2.629645, -0.800139, 1.570796, 2.190885],accel_mss,speed_ms,0,blend_radius_m)
  movel([0.618134, -1.286483, -2.627405, -0.798501, 1.570796, 2.188930],accel_mss,speed_ms,0,blend_radius_m)
  movel([0.615213, -1.290829, -2.624872, -0.796688, 1.570796, 2.186010],accel_mss,speed_ms,0,blend_radius_m)
  movel([0.611087, -1.295845, -2.621918, -0.794626, 1.570796, 2.181883],accel_mss,speed_ms,0,blend_radius_m)
  movel([0.607417, -1.299709, -2.619621, -0.793059, 1.570796, 2.178213],accel_mss,speed_ms,0,blend_radius_m)
  movel([0.603783, -1.303019, -2.617638, -0.791733, 1.570796, 2.174580],accel_mss,speed_ms,0,blend_radius_m)
  movel([0.600187, -1.305810, -2.615954, -0.790625, 1.570796, 2.170983],accel_mss,speed_ms,0,blend_radius_m)
  movel([0.596626, -1.308119, -2.614554, -0.789716, 1.570796, 2.167422],accel_mss,speed_ms,0,blend_radius_m)
  movel([0.593104, -1.309972, -2.613425, -0.788992, 1.570796, 2.163900],accel_mss,speed_ms,0,blend_radius_m)
  movel([0.589624, -1.311404, -2.612550, -0.788435, 1.570796, 2.160420],accel_mss,speed_ms,0,blend_radius_m)
  movel([0.586182, -1.312445, -2.611912, -0.788032, 1.570796, 2.156978],accel_mss,speed_ms,0,blend_radius_m)
  movel([0.582788, -1.313123, -2.611496, -0.787770, 1.570796, 2.153584],accel_mss,speed_ms,0,blend_radius_m)
  movel([0.579444, -1.313462, -2.611287, -0.787640, 1.570796, 2.150241],accel_mss,speed_ms,0,blend_radius_m)
  movel([0.576153, -1.313492, -2.611269, -0.787628, 1.570796, 2.146949],accel_mss,speed_ms,0,blend_radius_m)
  movel([0.569748, -1.312727, -2.611739, -0.787923, 1.570796, 2.140544],accel_mss,speed_ms,0,blend_radius_m)
  movel([0.563618, -1.311024, -2.612782, -0.788583, 1.570796, 2.134414],accel_mss,speed_ms,0,blend_radius_m)
  movel([0.557815, -1.308577, -2.614276, -0.789537, 1.570796, 2.128612],accel_mss,speed_ms,0,blend_radius_m)
  movel([0.552793, -1.305673, -2.616037, -0.790679, 1.570796, 2.123589],accel_mss,speed_ms,0,blend_radius_m)
  movel([0.546439, -1.301825, -2.618355, -0.792209, 1.570796, 2.117235],accel_mss,speed_ms,0,blend_radius_m)
  movel([0.538992, -1.298017, -2.620629, -0.793743, 1.570796, 2.109788],accel_mss,speed_ms,0,blend_radius_m)
  movel([0.534946, -1.296435, -2.621569, -0.794385, 1.570796, 2.105742],accel_mss,speed_ms,0,blend_radius_m)
  movel([0.530732, -1.295234, -2.622280, -0.794875, 1.570796, 2.101528],accel_mss,speed_ms,0,blend_radius_m)
  movel([0.526397, -1.294532, -2.622694, -0.795162, 1.570796, 2.097193],accel_mss,speed_ms,0,blend_radius_m)
  movel([0.521986, -1.294450, -2.622743, -0.795196, 1.570796, 2.092783],accel_mss,speed_ms,0,blend_radius_m)
  movel([0.517551, -1.295102, -2.622358, -0.794929, 1.570796, 2.088347],accel_mss,speed_ms,0,blend_radius_m)
  movel([0.513139, -1.296598, -2.621472, -0.794319, 1.570796, 2.083935],accel_mss,speed_ms,0,blend_radius_m)
  movel([0.510959, -1.297695, -2.620820, -0.793873, 1.570796, 2.081755],accel_mss,speed_ms,0,blend_radius_m)
  movel([0.508806, -1.299044, -2.620018, -0.793328, 1.570796, 2.079603],accel_mss,speed_ms,0,blend_radius_m)
  movel([0.506685, -1.300657, -2.619054, -0.792678, 1.570796, 2.077481],accel_mss,speed_ms,0,blend_radius_m)
  movel([0.504608, -1.302541, -2.617925, -0.791923, 1.570796, 2.075404],accel_mss,speed_ms,0,blend_radius_m)
  movel([0.502577, -1.304714, -2.616616, -0.791058, 1.570796, 2.073373],accel_mss,speed_ms,0,blend_radius_m)
  movel([0.500603, -1.307181, -2.615124, -0.790084, 1.570796, 2.071399],accel_mss,speed_ms,0,blend_radius_m)
  movel([0.496846, -1.313044, -2.611544, -0.787801, 1.570796, 2.067642],accel_mss,speed_ms,0,blend_radius_m)
  movel([0.495747, -1.315916, -2.609774, -0.786699, 1.570796, 2.066543],accel_mss,speed_ms,0,blend_radius_m)
  movel([0.495180, -1.318781, -2.607998, -0.785610, 1.570796, 2.065976],accel_mss,speed_ms,0,blend_radius_m)
  movel([0.495187, -1.321603, -2.606237, -0.784549, 1.570796, 2.065984],accel_mss,speed_ms,0,blend_radius_m)
  movel([0.495803, -1.324360, -2.604507, -0.783522, 1.570796, 2.066599],accel_mss,speed_ms,0,blend_radius_m)
  movel([0.498940, -1.320812, -2.606731, -0.784845, 1.570796, 2.069737],accel_mss,speed_ms,0,blend_radius_m)
  movel([0.502275, -1.317569, -2.608750, -0.786069, 1.570796, 2.073071],accel_mss,speed_ms,0,blend_radius_m)
  movel([0.505769, -1.314646, -2.610558, -0.787185, 1.570796, 2.076565],accel_mss,speed_ms,0,blend_radius_m)
  movel([0.509384, -1.312057, -2.612150, -0.788182, 1.570796, 2.080180],accel_mss,speed_ms,0,blend_radius_m)
  movel([0.513088, -1.309816, -2.613520, -0.789052, 1.570796, 2.083884],accel_mss,speed_ms,0,blend_radius_m)
  movel([0.516839, -1.307939, -2.614664, -0.789787, 1.570796, 2.087636],accel_mss,speed_ms,0,blend_radius_m)
  movel([0.520603, -1.306437, -2.615575, -0.790377, 1.570796, 2.091399],accel_mss,speed_ms,0,blend_radius_m)
  movel([0.524338, -1.305326, -2.616247, -0.790816, 1.570796, 2.095134],accel_mss,speed_ms,0,blend_radius_m)
  movel([0.528007, -1.304615, -2.616676, -0.791098, 1.570796, 2.098803],accel_mss,speed_ms,0,blend_radius_m)
  movel([0.531574, -1.304316, -2.616856, -0.791216, 1.570796, 2.102370],accel_mss,speed_ms,0,blend_radius_m)
  movel([0.534998, -1.304439, -2.616782, -0.791168, 1.570796, 2.105794],accel_mss,speed_ms,0,blend_radius_m)
  movel([0.538241, -1.304991, -2.616449, -0.790949, 1.570796, 2.109037],accel_mss,speed_ms,0,blend_radius_m)
  movel([0.541269, -1.305981, -2.615851, -0.790557, 1.570796, 2.112065],accel_mss,speed_ms,0,blend_radius_m)
  movel([0.544045, -1.307410, -2.614985, -0.789994, 1.570796, 2.114841],accel_mss,speed_ms,0,blend_radius_m)
  movel([0.546532, -1.309284, -2.613845, -0.789260, 1.570796, 2.117328],accel_mss,speed_ms,0,blend_radius_m)
  movel([0.548699, -1.311607, -2.612425, -0.788356, 1.570796, 2.119495],accel_mss,speed_ms,0,blend_radius_m)
  movel([0.550171, -1.313797, -2.611081, -0.787511, 1.570796, 2.120967],accel_mss,speed_ms,0,blend_radius_m)
  movel([0.551285, -1.316138, -2.609637, -0.786614, 1.570796, 2.122081],accel_mss,speed_ms,0,blend_radius_m)
  movel([0.552062, -1.318602, -2.608109, -0.785678, 1.570796, 2.122858],accel_mss,speed_ms,0,blend_radius_m)
  movel([0.552517, -1.321175, -2.606505, -0.784709, 1.570796, 2.123313],accel_mss,speed_ms,0,blend_radius_m)
  movel([0.552533, -1.326551, -2.603125, -0.782713, 1.570796, 2.123330],accel_mss,speed_ms,0,blend_radius_m)
  movel([0.551472, -1.332105, -2.599592, -0.780692, 1.570796, 2.122268],accel_mss,speed_ms,0,blend_radius_m)
  movel([0.549464, -1.337687, -2.596000, -0.778702, 1.570796, 2.120261],accel_mss,speed_ms,0,blend_radius_m)
  movel([0.546636, -1.343148, -2.592444, -0.776797, 1.570796, 2.117432],accel_mss,speed_ms,0,blend_radius_m)
  movel([0.543110, -1.348358, -2.589014, -0.775017, 1.570796, 2.113906],accel_mss,speed_ms,0,blend_radius_m)
  movel([0.538998, -1.353183, -2.585804, -0.773402, 1.570796, 2.109794],accel_mss,speed_ms,0,blend_radius_m)
  movel([0.534415, -1.357499, -2.582905, -0.771984, 1.570796, 2.105211],accel_mss,speed_ms,0,blend_radius_m)
  movel([0.529458, -1.361187, -2.580408, -0.770794, 1.570796, 2.100254],accel_mss,speed_ms,0,blend_radius_m)
  movel([0.524227, -1.364125, -2.578405, -0.769859, 1.570796, 2.095023],accel_mss,speed_ms,0,blend_radius_m)
  movel([0.521536, -1.365274, -2.577618, -0.769497, 1.570796, 2.092333],accel_mss,speed_ms,0,blend_radius_m)
  movel([0.518811, -1.366194, -2.576987, -0.769208, 1.570796, 2.089607],accel_mss,speed_ms,0,blend_radius_m)
  movel([0.516061, -1.366867, -2.576524, -0.768998, 1.570796, 2.086857],accel_mss,speed_ms,0,blend_radius_m)
  movel([0.513299, -1.367276, -2.576243, -0.768870, 1.570796, 2.084095],accel_mss,speed_ms,0,blend_radius_m)
  movel([0.510533, -1.367408, -2.576152, -0.768829, 1.570796, 2.081330],accel_mss,speed_ms,0,blend_radius_m)
  movel([0.507774, -1.367246, -2.576263, -0.768879, 1.570796, 2.078570],accel_mss,speed_ms,0,blend_radius_m)
  movel([0.505030, -1.366775, -2.576587, -0.769026, 1.570796, 2.075826],accel_mss,speed_ms,0,blend_radius_m)
  movel([0.502313, -1.365976, -2.577136, -0.769276, 1.570796, 2.073109],accel_mss,speed_ms,0,blend_radius_m)
  movel([0.499630, -1.364834, -2.577920, -0.769635, 1.570796, 2.070427],accel_mss,speed_ms,0,blend_radius_m)
  movel([0.496996, -1.363328, -2.578949, -0.770111, 1.570796, 2.067792],accel_mss,speed_ms,0,blend_radius_m)
  movel([0.495196, -1.361729, -2.580039, -0.770621, 1.570796, 2.065993],accel_mss,speed_ms,0,blend_radius_m)
  movel([0.490787, -1.356741, -2.583416, -0.772231, 1.570796, 2.061583],accel_mss,speed_ms,0,blend_radius_m)
  movel([0.488063, -1.352882, -2.586005, -0.773501, 1.570796, 2.058859],accel_mss,speed_ms,0,blend_radius_m)
  movel([0.485232, -1.348053, -2.589216, -0.775120, 1.570796, 2.056028],accel_mss,speed_ms,0,blend_radius_m)
  movel([0.482488, -1.342195, -2.593068, -0.777126, 1.570796, 2.053285],accel_mss,speed_ms,0,blend_radius_m)
  movel([0.480022, -1.335246, -2.597576, -0.779567, 1.570796, 2.050818],accel_mss,speed_ms,0,blend_radius_m)
  movel([0.478776, -1.330056, -2.600900, -0.781433, 1.570796, 2.049572],accel_mss,speed_ms,0,blend_radius_m)
  movel([0.478173, -1.325051, -2.604072, -0.783266, 1.570796, 2.048969],accel_mss,speed_ms,0,blend_radius_m)
  movel([0.478145, -1.320245, -2.607086, -0.785059, 1.570796, 2.048942],accel_mss,speed_ms,0,blend_radius_m)
  movel([0.478620, -1.315656, -2.609935, -0.786798, 1.570796, 2.049417],accel_mss,speed_ms,0,blend_radius_m)
  movel([0.479528, -1.311306, -2.612610, -0.788473, 1.570796, 2.050324],accel_mss,speed_ms,0,blend_radius_m)
  movel([0.480790, -1.307215, -2.615103, -0.790071, 1.570796, 2.051586],accel_mss,speed_ms,0,blend_radius_m)
  movel([0.482327, -1.303405, -2.617405, -0.791579, 1.570796, 2.053123],accel_mss,speed_ms,0,blend_radius_m)
  movel([0.484063, -1.299897, -2.619509, -0.792983, 1.570796, 2.054859],accel_mss,speed_ms,0,blend_radius_m)
  movel([0.487793, -1.293891, -2.623072, -0.795425, 1.570796, 2.058590],accel_mss,speed_ms,0,blend_radius_m)
  movel([0.491303, -1.289385, -2.625716, -0.797288, 1.570796, 2.062100],accel_mss,speed_ms,0,blend_radius_m)
  movel([0.493913, -1.286561, -2.627360, -0.798468, 1.570796, 2.064709],accel_mss,speed_ms,0,blend_radius_m)
  movel([0.494933, -1.285584, -2.627926, -0.798879, 1.570796, 2.065729],accel_mss,speed_ms,0,blend_radius_m)
  movel([0.499958, -1.281263, -2.630416, -0.800710, 1.570796, 2.070754],accel_mss,speed_ms,0,blend_radius_m)
  movel([0.504954, -1.277610, -2.632503, -0.802276, 1.570796, 2.075750],accel_mss,speed_ms,0,blend_radius_m)
  movel([0.509877, -1.274589, -2.634216, -0.803584, 1.570796, 2.080674],accel_mss,speed_ms,0,blend_radius_m)
  movel([0.514695, -1.272158, -2.635586, -0.804644, 1.570796, 2.085492],accel_mss,speed_ms,0,blend_radius_m)
  movel([0.519367, -1.270269, -2.636646, -0.805474, 1.570796, 2.090164],accel_mss,speed_ms,0,blend_radius_m)
  movel([0.523863, -1.268875, -2.637426, -0.806088, 1.570796, 2.094659],accel_mss,speed_ms,0,blend_radius_m)
  movel([0.528142, -1.267924, -2.637956, -0.806509, 1.570796, 2.098939],accel_mss,speed_ms,0,blend_radius_m)
  movel([0.532180, -1.267360, -2.638270, -0.806759, 1.570796, 2.102976],accel_mss,speed_ms,0,blend_radius_m)
  movel([0.539407, -1.267177, -2.638372, -0.806840, 1.570796, 2.110203],accel_mss,speed_ms,0,blend_radius_m)
  movel([0.545322, -1.267863, -2.637990, -0.806536, 1.570796, 2.116119],accel_mss,speed_ms,0,blend_radius_m)
  movel([0.549738, -1.268942, -2.637388, -0.806059, 1.570796, 2.120534],accel_mss,speed_ms,0,blend_radius_m)
  movel([0.552467, -1.269941, -2.636830, -0.805618, 1.570796, 2.123264],accel_mss,speed_ms,0,blend_radius_m)
  movel([0.558978, -1.272250, -2.635535, -0.804604, 1.570796, 2.129774],accel_mss,speed_ms,0,blend_radius_m)
  movel([0.565628, -1.275352, -2.633784, -0.803252, 1.570796, 2.136425],accel_mss,speed_ms,0,blend_radius_m)
  movel([0.572238, -1.278718, -2.631872, -0.801799, 1.570796, 2.143035],accel_mss,speed_ms,0,blend_radius_m)
  movel([0.578657, -1.281812, -2.630101, -0.800476, 1.570796, 2.149453],accel_mss,speed_ms,0,blend_radius_m)
  movel([0.584747, -1.284103, -2.628782, -0.799504, 1.570796, 2.155543],accel_mss,speed_ms,0,blend_radius_m)
  movel([0.587632, -1.284777, -2.628393, -0.799219, 1.570796, 2.158428],accel_mss,speed_ms,0,blend_radius_m)
  movel([0.590390, -1.285049, -2.628235, -0.799104, 1.570796, 2.161186],accel_mss,speed_ms,0,blend_radius_m)
  movel([0.593011, -1.284847, -2.628353, -0.799190, 1.570796, 2.163807],accel_mss,speed_ms,0,blend_radius_m)
  movel([0.595481, -1.284100, -2.628784, -0.799505, 1.570796, 2.166277],accel_mss,speed_ms,0,blend_radius_m)
  movel([0.597789, -1.282738, -2.629569, -0.800082, 1.570796, 2.168585],accel_mss,speed_ms,0,blend_radius_m)
  movel([0.599925, -1.280685, -2.630748, -0.800957, 1.570796, 2.170721],accel_mss,speed_ms,0,blend_radius_m)
  movel([0.601233, -1.278934, -2.631749, -0.801707, 1.570796, 2.172029],accel_mss,speed_ms,0,blend_radius_m)
  movel([0.602216, -1.277193, -2.632740, -0.802456, 1.570796, 2.173012],accel_mss,speed_ms,0,blend_radius_m)
  movel([0.603336, -1.273743, -2.634694, -0.803952, 1.570796, 2.174132],accel_mss,speed_ms,0,blend_radius_m)
  movel([0.603527, -1.270346, -2.636603, -0.805440, 1.570796, 2.174323],accel_mss,speed_ms,0,blend_radius_m)
  movel([0.603045, -1.267015, -2.638462, -0.806912, 1.570796, 2.173842],accel_mss,speed_ms,0,blend_radius_m)
  movel([0.601080, -1.260598, -2.642003, -0.809787, 1.570796, 2.171876],accel_mss,speed_ms,0,blend_radius_m)
  movel([0.600119, -1.257530, -2.643679, -0.811180, 1.570796, 2.170916],accel_mss,speed_ms,0,blend_radius_m)
  movel([0.599531, -1.254560, -2.645290, -0.812539, 1.570796, 2.170328],accel_mss,speed_ms,0,blend_radius_m)
  movel([0.599600, -1.249654, -2.647928, -0.814806, 1.570796, 2.170397],accel_mss,speed_ms,0,blend_radius_m)
  movel([0.600494, -1.243384, -2.651259, -0.817746, 1.570796, 2.171290],accel_mss,speed_ms,0,blend_radius_m)
  movel([0.602001, -1.236880, -2.654664, -0.820845, 1.570796, 2.172797],accel_mss,speed_ms,0,blend_radius_m)
  movel([0.603892, -1.231320, -2.657536, -0.823534, 1.570796, 2.174689],accel_mss,speed_ms,0,blend_radius_m)
  movel([0.605766, -1.227851, -2.659309, -0.825229, 1.570796, 2.176562],accel_mss,speed_ms,0,blend_radius_m)
  movel([0.608409, -1.223622, -2.661453, -0.827315, 1.570796, 2.179206],accel_mss,speed_ms,0,blend_radius_m)
  movel([0.610891, -1.219588, -2.663478, -0.829323, 1.570796, 2.181687],accel_mss,speed_ms,0,blend_radius_m)
  movel([0.612267, -1.216723, -2.664905, -0.830761, 1.570796, 2.183064],accel_mss,speed_ms,0,blend_radius_m)
  movel([0.612506, -1.213892, -2.666306, -0.832190, 1.570796, 2.183302],accel_mss,speed_ms,0,blend_radius_m)
  movel([0.612217, -1.210716, -2.667868, -0.833805, 1.570796, 2.183013],accel_mss,speed_ms,0,blend_radius_m)
  movel([0.611948, -1.207155, -2.669605, -0.835629, 1.570796, 2.182744],accel_mss,speed_ms,0,blend_radius_m)
  movel([0.612257, -1.203153, -2.671540, -0.837695, 1.570796, 2.183053],accel_mss,speed_ms,0,blend_radius_m)
  movel([0.613006, -1.200650, -2.672742, -0.838997, 1.570796, 2.183802],accel_mss,speed_ms,0,blend_radius_m)
  speed_ms = 0.003
  movel([0.613006, -1.193454, -2.669122, -0.849813, 1.570796, 2.183802],accel_mss,speed_ms,0,blend_radius_m)
  speed_ms = 0.01
  movel([0.613006, -1.166119, -2.654391, -0.891880, 1.570796, 2.183802],accel_mss,speed_ms,0,blend_radius_m)
  #M_RunCode9
  movel([0.480011, -1.274699, -2.598269, -0.839421, 1.570796, 2.050808],accel_mss,speed_ms,0,blend_radius_m)
  #M_RunCode3
  movel([0.480011, -1.300846, -2.611571, -0.799973, 1.570796, 2.050808],accel_mss,speed_ms,0,blend_radius_m)
  speed_ms = 0.003
  movel([0.480011, -1.307671, -2.614826, -0.789892, 1.570796, 2.050808],accel_mss,speed_ms,0,blend_radius_m)
  speed_ms = 0.007
  movel([0.473131, -1.306142, -2.615753, -0.790493, 1.570796, 2.043927],accel_mss,speed_ms,0,blend_radius_m)
  movel([0.466158, -1.305516, -2.616132, -0.790741, 1.570796, 2.036954],accel_mss,speed_ms,0,blend_radius_m)
  movel([0.459184, -1.305685, -2.616030, -0.790674, 1.570796, 2.029980],accel_mss,speed_ms,0,blend_radius_m)
  movel([0.452290, -1.306536, -2.615515, -0.790338, 1.570796, 2.023086],accel_mss,speed_ms,0,blend_radius_m)
  movel([0.445562, -1.307953, -2.614655, -0.789781, 1.570796, 2.016358],accel_mss,speed_ms,0,blend_radius_m)
  movel([0.439080, -1.309822, -2.613517, -0.789050, 1.570796, 2.009876],accel_mss,speed_ms,0,blend_radius_m)
  movel([0.432919, -1.312027, -2.612168, -0.788194, 1.570796, 2.003715],accel_mss,speed_ms,0,blend_radius_m)
  movel([0.427145, -1.314454, -2.610676, -0.787258, 1.570796, 1.997942],accel_mss,speed_ms,0,blend_radius_m)
  movel([0.421831, -1.316991, -2.609109, -0.786289, 1.570796, 1.992627],accel_mss,speed_ms,0,blend_radius_m)
  movel([0.417038, -1.319526, -2.607534, -0.785329, 1.570796, 1.987835],accel_mss,speed_ms,0,blend_radius_m)
  movel([0.409259, -1.324170, -2.604626, -0.783592, 1.570796, 1.980055],accel_mss,speed_ms,0,blend_radius_m)
  movel([0.404262, -1.327550, -2.602493, -0.782347, 1.570796, 1.975059],accel_mss,speed_ms,0,blend_radius_m)
  movel([0.402496, -1.328854, -2.601665, -0.781870, 1.570796, 1.973292],accel_mss,speed_ms,0,blend_radius_m)
  movel([0.399641, -1.330838, -2.600402, -0.781149, 1.570796, 1.970437],accel_mss,speed_ms,0,blend_radius_m)
  movel([0.392413, -1.336510, -2.596761, -0.779118, 1.570796, 1.963210],accel_mss,speed_ms,0,blend_radius_m)
  movel([0.387795, -1.340589, -2.594116, -0.777685, 1.570796, 1.958592],accel_mss,speed_ms,0,blend_radius_m)
  movel([0.382850, -1.345411, -2.590959, -0.776019, 1.570796, 1.953646],accel_mss,speed_ms,0,blend_radius_m)
  movel([0.377828, -1.350912, -2.587319, -0.774158, 1.570796, 1.948624],accel_mss,speed_ms,0,blend_radius_m)
  movel([0.372976, -1.357023, -2.583227, -0.772140, 1.570796, 1.943773],accel_mss,speed_ms,0,blend_radius_m)
  movel([0.368538, -1.363669, -2.578717, -0.770004, 1.570796, 1.939335],accel_mss,speed_ms,0,blend_radius_m)
  movel([0.364744, -1.370784, -2.573819, -0.767785, 1.570796, 1.935541],accel_mss,speed_ms,0,blend_radius_m)
  movel([0.363161, -1.374498, -2.571235, -0.766656, 1.570796, 1.933957],accel_mss,speed_ms,0,blend_radius_m)
  movel([0.361821, -1.378304, -2.568566, -0.765519, 1.570796, 1.932617],accel_mss,speed_ms,0,blend_radius_m)
  movel([0.360750, -1.382195, -2.565816, -0.764378, 1.570796, 1.931546],accel_mss,speed_ms,0,blend_radius_m)
  movel([0.359975, -1.386165, -2.562988, -0.763236, 1.570796, 1.930771],accel_mss,speed_ms,0,blend_radius_m)
  movel([0.359520, -1.390207, -2.560085, -0.762097, 1.570796, 1.930317],accel_mss,speed_ms,0,blend_radius_m)
  movel([0.359411, -1.394315, -2.557111, -0.760963, 1.570796, 1.930207],accel_mss,speed_ms,0,blend_radius_m)
  movel([0.359669, -1.398483, -2.554068, -0.759838, 1.570796, 1.930465],accel_mss,speed_ms,0,blend_radius_m)
  movel([0.360313, -1.402708, -2.550958, -0.758724, 1.570796, 1.931109],accel_mss,speed_ms,0,blend_radius_m)
  movel([0.361370, -1.406985, -2.547782, -0.757622, 1.570796, 1.932166],accel_mss,speed_ms,0,blend_radius_m)
  movel([0.362857, -1.411313, -2.544541, -0.756534, 1.570796, 1.933653],accel_mss,speed_ms,0,blend_radius_m)
  movel([0.364793, -1.415688, -2.541238, -0.755463, 1.570796, 1.935590],accel_mss,speed_ms,0,blend_radius_m)
  movel([0.367197, -1.420112, -2.537868, -0.754409, 1.570796, 1.937994],accel_mss,speed_ms,0,blend_radius_m)
  movel([0.367412, -1.420438, -2.537619, -0.754332, 1.570796, 1.938209],accel_mss,speed_ms,0,blend_radius_m)
  movel([0.370499, -1.424346, -2.534616, -0.753427, 1.570796, 1.941296],accel_mss,speed_ms,0,blend_radius_m)
  movel([0.373678, -1.427760, -2.531974, -0.752655, 1.570796, 1.944475],accel_mss,speed_ms,0,blend_radius_m)
  movel([0.376936, -1.430712, -2.529675, -0.752002, 1.570796, 1.947732],accel_mss,speed_ms,0,blend_radius_m)
  movel([0.380264, -1.433229, -2.527705, -0.751455, 1.570796, 1.951060],accel_mss,speed_ms,0,blend_radius_m)
  movel([0.383650, -1.435340, -2.526046, -0.751003, 1.570796, 1.954446],accel_mss,speed_ms,0,blend_radius_m)
  movel([0.387084, -1.437071, -2.524679, -0.750638, 1.570796, 1.957881],accel_mss,speed_ms,0,blend_radius_m)
  movel([0.390559, -1.438445, -2.523592, -0.750352, 1.570796, 1.961355],accel_mss,speed_ms,0,blend_radius_m)
  movel([0.394061, -1.439489, -2.522764, -0.750136, 1.570796, 1.964857],accel_mss,speed_ms,0,blend_radius_m)
  movel([0.397580, -1.440229, -2.522176, -0.749984, 1.570796, 1.968376],accel_mss,speed_ms,0,blend_radius_m)
  movel([0.401104, -1.440683, -2.521814, -0.749891, 1.570796, 1.971901],accel_mss,speed_ms,0,blend_radius_m)
  movel([0.404624, -1.440877, -2.521660, -0.749852, 1.570796, 1.975421],accel_mss,speed_ms,0,blend_radius_m)
  movel([0.408127, -1.440833, -2.521695, -0.749861, 1.570796, 1.978923],accel_mss,speed_ms,0,blend_radius_m)
  movel([0.415037, -1.440122, -2.522261, -0.750006, 1.570796, 1.985833],accel_mss,speed_ms,0,blend_radius_m)
  movel([0.421731, -1.438723, -2.523371, -0.750294, 1.570796, 1.992527],accel_mss,speed_ms,0,blend_radius_m)
  movel([0.428105, -1.436813, -2.524883, -0.750692, 1.570796, 1.998901],accel_mss,speed_ms,0,blend_radius_m)
  movel([0.434046, -1.434567, -2.526654, -0.751168, 1.570796, 2.004842],accel_mss,speed_ms,0,blend_radius_m)
  movel([0.439434, -1.432158, -2.528545, -0.751686, 1.570796, 2.010230],accel_mss,speed_ms,0,blend_radius_m)
  movel([0.444144, -1.429770, -2.530410, -0.752209, 1.570796, 2.014940],accel_mss,speed_ms,0,blend_radius_m)
  movel([0.450999, -1.425793, -2.533498, -0.753098, 1.570796, 2.021796],accel_mss,speed_ms,0,blend_radius_m)
  movel([0.453527, -1.424126, -2.534785, -0.753478, 1.570796, 2.024324],accel_mss,speed_ms,0,blend_radius_m)
  movel([0.455076, -1.423162, -2.535528, -0.753699, 1.570796, 2.025872],accel_mss,speed_ms,0,blend_radius_m)
  movel([0.459274, -1.420318, -2.537711, -0.754361, 1.570796, 2.030070],accel_mss,speed_ms,0,blend_radius_m)
  movel([0.465446, -1.415673, -2.541249, -0.755467, 1.570796, 2.036242],accel_mss,speed_ms,0,blend_radius_m)
  movel([0.472944, -1.409280, -2.546067, -0.757042, 1.570796, 2.043740],accel_mss,speed_ms,0,blend_radius_m)
  movel([0.476985, -1.405440, -2.548932, -0.758017, 1.570796, 2.047781],accel_mss,speed_ms,0,blend_radius_m)
  movel([0.481113, -1.401173, -2.552091, -0.759126, 1.570796, 2.051909],accel_mss,speed_ms,0,blend_radius_m)
  movel([0.485244, -1.396479, -2.555534, -0.760376, 1.570796, 2.056040],accel_mss,speed_ms,0,blend_radius_m)
  movel([0.489291, -1.391359, -2.559253, -0.761777, 1.570796, 2.060088],accel_mss,speed_ms,0,blend_radius_m)
  movel([0.493170, -1.385810, -2.563242, -0.763337, 1.570796, 2.063967],accel_mss,speed_ms,0,blend_radius_m)
  movel([0.496793, -1.379827, -2.567492, -0.765070, 1.570796, 2.067589],accel_mss,speed_ms,0,blend_radius_m)
  movel([0.500067, -1.373407, -2.571996, -0.766986, 1.570796, 2.070863],accel_mss,speed_ms,0,blend_radius_m)
  movel([0.502898, -1.366546, -2.576745, -0.769098, 1.570796, 2.073695],accel_mss,speed_ms,0,blend_radius_m)
  speed_ms = 0.003
  movel([0.502898, -1.359997, -2.573686, -0.778706, 1.570796, 2.073695],accel_mss,speed_ms,0,blend_radius_m)
  speed_ms = 0.01
  movel([0.502898, -1.334806, -2.561165, -0.816418, 1.570796, 2.073695],accel_mss,speed_ms,0,blend_radius_m)
  #M_RunCode9
  movel([0.474292, -1.328447, -2.565310, -0.818632, 1.570796, 2.045088],accel_mss,speed_ms,0,blend_radius_m)
  #M_RunCode3
